Universal Robots URScript: test_first_drawing_6.script

def Machining1():
  # Default parameters:
  global speed_ms = 0.3
  global speed_rads = 0.75
  global accel_mss = 3
  global accel_radss = 1.2
  global blend_radius_m = 0.001

  # Add subprograms here
  # Start of main program
  # Program generated by RoboDK v5.6.5 for UR10e on 02/02/2024 17:00:01
  # Using nominal kinematics.
  blend_radius_m = 0.001
  speed_ms = 1.000
  # set_reference(p[0.133734, -0.230000, -0.011586, 0.000000, 0.000000, 0.000000])
  set_tcp(p[0.000000, 0.000000, 0.252000, 0.000000, 0.000000, 0.000000])
  # Show Tool
  movej([-0.330517, -0.652308, -2.595548, -1.464533, 1.570796, 1.240279],accel_radss,speed_rads,0,blend_radius_m)
  movel([-0.330517, -0.652308, -2.595548, -1.464533, 1.570796, 1.240279],accel_mss,speed_ms,0,blend_radius_m)
  # Splitting Linear movement in 6 (instruction 7: MoveL 3)
  movel([-0.330517, -0.658933, -2.623995, -1.429460, 1.570796, 1.240279],accel_mss,speed_ms,0,blend_radius_m)
  movel([-0.330517, -0.667915, -2.652250, -1.392224, 1.570796, 1.240279],accel_mss,speed_ms,0,blend_radius_m)
  movel([-0.330517, -0.679637, -2.680305, -1.352447, 1.570796, 1.240279],accel_mss,speed_ms,0,blend_radius_m)
  movel([-0.330517, -0.694570, -2.708148, -1.309671, 1.570796, 1.240279],accel_mss,speed_ms,0,blend_radius_m)
  movel([-0.330517, -0.713300, -2.735763, -1.263326, 1.570796, 1.240279],accel_mss,speed_ms,0,blend_radius_m)
  movel([-0.330517, -0.736556, -2.763126, -1.212708, 1.570796, 1.240279],accel_mss,speed_ms,0,blend_radius_m)
  movel([-0.330517, -0.736556, -2.763126, -1.212708, 1.570796, 1.240279],accel_mss,speed_ms,0,blend_radius_m)
  speed_ms = 1.000
  movel([-0.330517, -0.736556, -2.763126, -1.212708, 1.570796, 1.240279],accel_mss,speed_ms,0,blend_radius_m)
  movel([-0.330517, -0.736556, -2.763126, -1.212708, 1.570796, 1.240279],accel_mss,speed_ms,0,blend_radius_m)
  movel([-0.330517, -0.736556, -2.763126, -1.212708, 1.570796, 1.240279],accel_mss,speed_ms,0,blend_radius_m)
  speed_ms = 0.005
  movel([-0.330517, -0.709218, -2.730259, -1.272912, 1.570796, 1.240279],accel_mss,speed_ms,0,blend_radius_m)
  speed_ms = 1.000
  movel([-0.330517, -0.736556, -2.763126, -1.212708, 1.570796, 1.240279],accel_mss,speed_ms,0,blend_radius_m)
  speed_ms = 0.040
  movel([-0.330517, -0.736556, -2.763126, -1.212708, 1.570796, 1.240279],accel_mss,speed_ms,0,blend_radius_m)
  speed_ms = 1.000
  movel([-0.330517, -0.736556, -2.763126, -1.212708, 1.570796, 1.240279],accel_mss,speed_ms,0,blend_radius_m)
  # Splitting Linear movement in 8 (instruction 21: MoveL 12)
  movel([-0.265752, -0.726906, -2.764568, -1.220915, 1.570796, 1.305044],accel_mss,speed_ms,0,blend_radius_m)
  movel([-0.203429, -0.722340, -2.765235, -1.224814, 1.570796, 1.367367],accel_mss,speed_ms,0,blend_radius_m)
  movel([-0.144075, -0.722992, -2.765140, -1.224257, 1.570796, 1.426722],accel_mss,speed_ms,0,blend_radius_m)
  movel([-0.088098, -0.728842, -2.764283, -1.219264, 1.570796, 1.482698],accel_mss,speed_ms,0,blend_radius_m)
  movel([-0.035774, -0.739721, -2.762642, -1.210026, 1.570796, 1.535022],accel_mss,speed_ms,0,blend_radius_m)
  movel([0.012756, -0.755321, -2.760186, -1.196882, 1.570796, 1.583552],accel_mss,speed_ms,0,blend_radius_m)
  movel([0.057475, -0.775222, -2.756871, -1.180296, 1.570796, 1.628271],accel_mss,speed_ms,0,blend_radius_m)
  movel([0.098470, -0.798920, -2.752649, -1.160820, 1.570796, 1.669266],accel_mss,speed_ms,0,blend_radius_m)
  speed_ms = 0.005
  movel([0.098470, -0.837473, -2.784197, -1.090719, 1.570796, 1.669266],accel_mss,speed_ms,0,blend_radius_m)
  speed_ms = 0.025
  movel([0.094484, -0.848078, -2.782141, -1.082170, 1.570796, 1.665281],accel_mss,speed_ms,0,blend_radius_m)
  movel([0.092287, -0.853406, -2.781085, -1.077898, 1.570796, 1.663083],accel_mss,speed_ms,0,blend_radius_m)
  movel([0.089913, -0.858734, -2.780012, -1.073643, 1.570796, 1.660710],accel_mss,speed_ms,0,blend_radius_m)
  movel([0.087338, -0.864042, -2.778926, -1.069420, 1.570796, 1.658135],accel_mss,speed_ms,0,blend_radius_m)
  movel([0.084536, -0.869315, -2.777832, -1.065242, 1.570796, 1.655333],accel_mss,speed_ms,0,blend_radius_m)
  movel([0.081477, -0.874542, -2.776731, -1.061116, 1.570796, 1.652273],accel_mss,speed_ms,0,blend_radius_m)
  movel([0.078131, -0.879702, -2.775628, -1.057059, 1.570796, 1.648928],accel_mss,speed_ms,0,blend_radius_m)
  movel([0.079373, -0.877446, -2.776112, -1.058831, 1.570796, 1.650169],accel_mss,speed_ms,0,blend_radius_m)
  movel([0.080517, -0.874618, -2.776715, -1.061056, 1.570796, 1.651313],accel_mss,speed_ms,0,blend_radius_m)
  movel([0.081210, -0.871968, -2.777275, -1.063146, 1.570796, 1.652007],accel_mss,speed_ms,0,blend_radius_m)
  movel([0.081271, -0.870953, -2.777489, -1.063947, 1.570796, 1.652068],accel_mss,speed_ms,0,blend_radius_m)
  movel([0.081086, -0.870269, -2.777632, -1.064488, 1.570796, 1.651882],accel_mss,speed_ms,0,blend_radius_m)
  movel([0.080605, -0.869994, -2.777690, -1.064705, 1.570796, 1.651401],accel_mss,speed_ms,0,blend_radius_m)
  movel([0.079917, -0.870224, -2.777642, -1.064524, 1.570796, 1.650713],accel_mss,speed_ms,0,blend_radius_m)
  movel([0.079063, -0.870887, -2.777502, -1.063999, 1.570796, 1.649859],accel_mss,speed_ms,0,blend_radius_m)
  movel([0.078060, -0.871934, -2.777282, -1.063173, 1.570796, 1.648856],accel_mss,speed_ms,0,blend_radius_m)
  movel([0.075754, -0.874898, -2.776655, -1.060835, 1.570796, 1.646551],accel_mss,speed_ms,0,blend_radius_m)
  movel([0.073242, -0.878610, -2.775863, -1.057916, 1.570796, 1.644038],accel_mss,speed_ms,0,blend_radius_m)
  movel([0.068514, -0.886327, -2.774188, -1.051873, 1.570796, 1.639311],accel_mss,speed_ms,0,blend_radius_m)
  movel([0.065663, -0.891230, -2.773106, -1.048053, 1.570796, 1.636460],accel_mss,speed_ms,0,blend_radius_m)
  movel([0.061416, -0.898083, -2.771568, -1.042738, 1.570796, 1.632212],accel_mss,speed_ms,0,blend_radius_m)
  movel([0.059067, -0.901365, -2.770821, -1.040203, 1.570796, 1.629863],accel_mss,speed_ms,0,blend_radius_m)
  movel([0.056470, -0.904440, -2.770115, -1.037833, 1.570796, 1.627267],accel_mss,speed_ms,0,blend_radius_m)
  movel([0.057008, -0.903519, -2.770327, -1.038543, 1.570796, 1.627804],accel_mss,speed_ms,0,blend_radius_m)
  movel([0.057386, -0.902191, -2.770632, -1.039565, 1.570796, 1.628182],accel_mss,speed_ms,0,blend_radius_m)
  movel([0.057710, -0.898919, -2.771378, -1.042091, 1.570796, 1.628506],accel_mss,speed_ms,0,blend_radius_m)
  movel([0.057532, -0.895865, -2.772069, -1.044455, 1.570796, 1.628328],accel_mss,speed_ms,0,blend_radius_m)
  movel([0.057276, -0.894808, -2.772307, -1.045274, 1.570796, 1.628072],accel_mss,speed_ms,0,blend_radius_m)
  movel([0.056930, -0.894278, -2.772426, -1.045686, 1.570796, 1.627726],accel_mss,speed_ms,0,blend_radius_m)
  movel([0.055907, -0.894028, -2.772481, -1.045879, 1.570796, 1.626704],accel_mss,speed_ms,0,blend_radius_m)
  movel([0.054873, -0.894325, -2.772415, -1.045649, 1.570796, 1.625669],accel_mss,speed_ms,0,blend_radius_m)
  movel([0.053834, -0.895056, -2.772251, -1.045082, 1.570796, 1.624631],accel_mss,speed_ms,0,blend_radius_m)
  movel([0.052803, -0.896120, -2.772012, -1.044258, 1.570796, 1.623599],accel_mss,speed_ms,0,blend_radius_m)
  movel([0.050825, -0.898766, -2.771413, -1.042210, 1.570796, 1.621621],accel_mss,speed_ms,0,blend_radius_m)
  movel([0.049035, -0.901386, -2.770816, -1.040187, 1.570796, 1.619831],accel_mss,speed_ms,0,blend_radius_m)
  movel([0.046096, -0.905333, -2.769909, -1.037147, 1.570796, 1.616892],accel_mss,speed_ms,0,blend_radius_m)
  movel([0.043104, -0.908938, -2.769072, -1.034379, 1.570796, 1.613900],accel_mss,speed_ms,0,blend_radius_m)
  movel([0.039882, -0.912201, -2.768307, -1.031881, 1.570796, 1.610679],accel_mss,speed_ms,0,blend_radius_m)
  movel([0.036270, -0.915096, -2.767623, -1.029670, 1.570796, 1.607066],accel_mss,speed_ms,0,blend_radius_m)
  movel([0.038295, -0.912091, -2.768333, -1.031965, 1.570796, 1.609092],accel_mss,speed_ms,0,blend_radius_m)
  movel([0.039935, -0.909052, -2.769046, -1.034292, 1.570796, 1.610731],accel_mss,speed_ms,0,blend_radius_m)
  movel([0.040448, -0.907548, -2.769396, -1.035445, 1.570796, 1.611244],accel_mss,speed_ms,0,blend_radius_m)
  movel([0.040644, -0.906186, -2.769712, -1.036491, 1.570796, 1.611440],accel_mss,speed_ms,0,blend_radius_m)
  movel([0.040480, -0.905086, -2.769966, -1.037336, 1.570796, 1.611276],accel_mss,speed_ms,0,blend_radius_m)
  movel([0.039889, -0.904398, -2.770125, -1.037866, 1.570796, 1.610686],accel_mss,speed_ms,0,blend_radius_m)
  movel([0.038611, -0.904273, -2.770154, -1.037962, 1.570796, 1.609407],accel_mss,speed_ms,0,blend_radius_m)
  movel([0.036998, -0.904844, -2.770022, -1.037523, 1.570796, 1.607794],accel_mss,speed_ms,0,blend_radius_m)
  movel([0.035210, -0.905879, -2.769783, -1.036727, 1.570796, 1.606006],accel_mss,speed_ms,0,blend_radius_m)
  movel([0.033415, -0.907124, -2.769494, -1.035771, 1.570796, 1.604211],accel_mss,speed_ms,0,blend_radius_m)
  speed_ms = 0.005
  movel([0.033415, -0.898152, -2.763466, -1.050771, 1.570796, 1.604211],accel_mss,speed_ms,0,blend_radius_m)
  speed_ms = 0.040
  movel([0.037572, -0.930926, -2.755578, -1.025884, 1.570796, 1.608368],accel_mss,speed_ms,0,blend_radius_m)
  speed_ms = 0.005
  movel([0.037572, -0.940094, -2.761488, -1.010807, 1.570796, 1.608368],accel_mss,speed_ms,0,blend_radius_m)
  speed_ms = 0.025
  movel([0.038407, -0.937648, -2.762106, -1.012634, 1.570796, 1.609204],accel_mss,speed_ms,0,blend_radius_m)
  movel([0.039504, -0.935133, -2.762738, -1.014518, 1.570796, 1.610300],accel_mss,speed_ms,0,blend_radius_m)
  movel([0.040832, -0.932593, -2.763372, -1.016424, 1.570796, 1.611628],accel_mss,speed_ms,0,blend_radius_m)
  movel([0.042377, -0.930056, -2.764001, -1.018332, 1.570796, 1.613173],accel_mss,speed_ms,0,blend_radius_m)
  movel([0.044112, -0.927559, -2.764616, -1.020214, 1.570796, 1.614908],accel_mss,speed_ms,0,blend_radius_m)
  movel([0.046017, -0.925143, -2.765207, -1.022039, 1.570796, 1.616813],accel_mss,speed_ms,0,blend_radius_m)
  movel([0.048065, -0.922844, -2.765765, -1.023780, 1.570796, 1.618862],accel_mss,speed_ms,0,blend_radius_m)
  movel([0.050239, -0.920694, -2.766285, -1.025410, 1.570796, 1.621035],accel_mss,speed_ms,0,blend_radius_m)
  movel([0.053602, -0.917840, -2.766970, -1.027579, 1.570796, 1.624398],accel_mss,speed_ms,0,blend_radius_m)
  movel([0.056890, -0.915555, -2.767514, -1.029320, 1.570796, 1.627686],accel_mss,speed_ms,0,blend_radius_m)
  movel([0.060092, -0.913802, -2.767930, -1.030657, 1.570796, 1.630888],accel_mss,speed_ms,0,blend_radius_m)
  movel([0.063188, -0.912552, -2.768225, -1.031612, 1.570796, 1.633984],accel_mss,speed_ms,0,blend_radius_m)
  movel([0.066168, -0.911768, -2.768409, -1.032211, 1.570796, 1.636964],accel_mss,speed_ms,0,blend_radius_m)
  movel([0.069022, -0.911415, -2.768492, -1.032482, 1.570796, 1.639818],accel_mss,speed_ms,0,blend_radius_m)
  movel([0.071734, -0.911461, -2.768482, -1.032447, 1.570796, 1.642530],accel_mss,speed_ms,0,blend_radius_m)
  movel([0.074296, -0.911861, -2.768387, -1.032140, 1.570796, 1.645092],accel_mss,speed_ms,0,blend_radius_m)
  movel([0.076697, -0.912580, -2.768218, -1.031591, 1.570796, 1.647493],accel_mss,speed_ms,0,blend_radius_m)
  movel([0.078931, -0.913578, -2.767983, -1.030829, 1.570796, 1.649727],accel_mss,speed_ms,0,blend_radius_m)
  movel([0.082865, -0.916242, -2.767351, -1.028797, 1.570796, 1.653661],accel_mss,speed_ms,0,blend_radius_m)
  movel([0.086044, -0.919518, -2.766568, -1.026304, 1.570796, 1.656840],accel_mss,speed_ms,0,blend_radius_m)
  movel([0.088410, -0.923091, -2.765706, -1.023593, 1.570796, 1.659206],accel_mss,speed_ms,0,blend_radius_m)
  movel([0.090331, -0.927270, -2.764687, -1.020432, 1.570796, 1.661127],accel_mss,speed_ms,0,blend_radius_m)
  movel([0.091833, -0.931808, -2.763567, -1.017014, 1.570796, 1.662629],accel_mss,speed_ms,0,blend_radius_m)
  movel([0.092966, -0.936641, -2.762360, -1.013388, 1.570796, 1.663762],accel_mss,speed_ms,0,blend_radius_m)
  movel([0.093774, -0.941716, -2.761075, -1.009597, 1.570796, 1.664570],accel_mss,speed_ms,0,blend_radius_m)
  movel([0.094306, -0.946974, -2.759726, -1.005688, 1.570796, 1.665103],accel_mss,speed_ms,0,blend_radius_m)
  movel([0.094614, -0.952360, -2.758325, -1.001704, 1.570796, 1.665411],accel_mss,speed_ms,0,blend_radius_m)
  movel([0.094736, -0.963302, -2.755416, -0.993671, 1.570796, 1.665532],accel_mss,speed_ms,0,blend_radius_m)
  movel([0.094750, -0.970923, -2.753340, -0.988126, 1.570796, 1.665546],accel_mss,speed_ms,0,blend_radius_m)
  movel([0.095064, -0.974489, -2.752355, -0.985545, 1.570796, 1.665861],accel_mss,speed_ms,0,blend_radius_m)
  movel([0.095787, -0.977736, -2.751449, -0.983203, 1.570796, 1.666583],accel_mss,speed_ms,0,blend_radius_m)
  movel([0.097346, -0.981517, -2.750386, -0.980486, 1.570796, 1.668143],accel_mss,speed_ms,0,blend_radius_m)
  movel([0.098905, -0.985307, -2.749309, -0.977773, 1.570796, 1.669701],accel_mss,speed_ms,0,blend_radius_m)
  movel([0.099406, -0.987343, -2.748726, -0.976320, 1.570796, 1.670202],accel_mss,speed_ms,0,blend_radius_m)
  movel([0.099571, -0.989546, -2.748092, -0.974750, 1.570796, 1.670367],accel_mss,speed_ms,0,blend_radius_m)
  movel([0.099295, -0.991964, -2.747392, -0.973033, 1.570796, 1.670091],accel_mss,speed_ms,0,blend_radius_m)
  movel([0.098473, -0.994652, -2.746609, -0.971128, 1.570796, 1.669269],accel_mss,speed_ms,0,blend_radius_m)
  movel([0.101094, -0.987874, -2.748574, -0.975941, 1.570796, 1.671890],accel_mss,speed_ms,0,blend_radius_m)
  movel([0.103419, -0.981143, -2.750492, -0.980754, 1.570796, 1.674215],accel_mss,speed_ms,0,blend_radius_m)
  movel([0.107547, -0.967644, -2.754238, -0.990506, 1.570796, 1.678343],accel_mss,speed_ms,0,blend_radius_m)
  movel([0.109649, -0.960093, -2.756278, -0.996019, 1.570796, 1.680446],accel_mss,speed_ms,0,blend_radius_m)
  movel([0.111578, -0.952541, -2.758278, -1.001571, 1.570796, 1.682375],accel_mss,speed_ms,0,blend_radius_m)
  movel([0.115043, -0.937387, -2.762172, -1.012830, 1.570796, 1.685839],accel_mss,speed_ms,0,blend_radius_m)
  movel([0.118016, -0.922483, -2.765853, -1.024053, 1.570796, 1.688812],accel_mss,speed_ms,0,blend_radius_m)
  movel([0.119175, -0.915076, -2.767628, -1.029685, 1.570796, 1.689972],accel_mss,speed_ms,0,blend_radius_m)
  movel([0.119952, -0.907871, -2.769321, -1.035197, 1.570796, 1.690749],accel_mss,speed_ms,0,blend_radius_m)
  movel([0.120167, -0.902405, -2.770583, -1.039401, 1.570796, 1.690963],accel_mss,speed_ms,0,blend_radius_m)
  movel([0.120127, -0.897049, -2.771802, -1.043538, 1.570796, 1.690923],accel_mss,speed_ms,0,blend_radius_m)
  movel([0.120107, -0.891619, -2.773019, -1.047751, 1.570796, 1.690904],accel_mss,speed_ms,0,blend_radius_m)
  movel([0.120387, -0.885931, -2.774275, -1.052183, 1.570796, 1.691183],accel_mss,speed_ms,0,blend_radius_m)
  movel([0.120647, -0.884307, -2.774630, -1.053451, 1.570796, 1.691443],accel_mss,speed_ms,0,blend_radius_m)
  movel([0.121203, -0.882545, -2.775013, -1.054830, 1.570796, 1.692000],accel_mss,speed_ms,0,blend_radius_m)
  movel([0.122110, -0.880885, -2.775373, -1.056131, 1.570796, 1.692906],accel_mss,speed_ms,0,blend_radius_m)
  movel([0.122719, -0.880160, -2.775529, -1.056700, 1.570796, 1.693515],accel_mss,speed_ms,0,blend_radius_m)
  movel([0.123441, -0.879540, -2.775663, -1.057186, 1.570796, 1.694238],accel_mss,speed_ms,0,blend_radius_m)
  movel([0.124465, -0.879007, -2.775777, -1.057605, 1.570796, 1.695262],accel_mss,speed_ms,0,blend_radius_m)
  movel([0.125422, -0.878749, -2.775833, -1.057807, 1.570796, 1.696219],accel_mss,speed_ms,0,blend_radius_m)
  movel([0.130425, -0.878041, -2.775985, -1.058363, 1.570796, 1.701221],accel_mss,speed_ms,0,blend_radius_m)
  movel([0.134885, -0.878093, -2.775974, -1.058323, 1.570796, 1.705681],accel_mss,speed_ms,0,blend_radius_m)
  movel([0.138838, -0.878832, -2.775815, -1.057742, 1.570796, 1.709634],accel_mss,speed_ms,0,blend_radius_m)
  movel([0.142320, -0.880210, -2.775519, -1.056661, 1.570796, 1.713117],accel_mss,speed_ms,0,blend_radius_m)
  movel([0.145368, -0.882154, -2.775098, -1.055137, 1.570796, 1.716164],accel_mss,speed_ms,0,blend_radius_m)
  movel([0.148021, -0.884600, -2.774566, -1.053223, 1.570796, 1.718817],accel_mss,speed_ms,0,blend_radius_m)
  movel([0.150317, -0.887485, -2.773934, -1.050970, 1.570796, 1.721113],accel_mss,speed_ms,0,blend_radius_m)
  movel([0.152293, -0.890749, -2.773213, -1.048427, 1.570796, 1.723089],accel_mss,speed_ms,0,blend_radius_m)
  movel([0.153993, -0.894325, -2.772415, -1.045649, 1.570796, 1.724789],accel_mss,speed_ms,0,blend_radius_m)
  movel([0.155459, -0.898148, -2.771553, -1.042688, 1.570796, 1.726255],accel_mss,speed_ms,0,blend_radius_m)
  movel([0.157842, -0.906294, -2.769687, -1.036408, 1.570796, 1.728639],accel_mss,speed_ms,0,blend_radius_m)
  movel([0.161526, -0.922971, -2.765735, -1.023684, 1.570796, 1.732322],accel_mss,speed_ms,0,blend_radius_m)
  movel([0.162250, -0.925447, -2.765132, -1.021810, 1.570796, 1.733046],accel_mss,speed_ms,0,blend_radius_m)
  movel([0.162856, -0.926430, -2.764892, -1.021067, 1.570796, 1.733653],accel_mss,speed_ms,0,blend_radius_m)
  movel([0.163731, -0.927104, -2.764727, -1.020558, 1.570796, 1.734527],accel_mss,speed_ms,0,blend_radius_m)
  movel([0.165528, -0.927367, -2.764663, -1.020359, 1.570796, 1.736325],accel_mss,speed_ms,0,blend_radius_m)
  movel([0.166517, -0.927169, -2.764711, -1.020509, 1.570796, 1.737313],accel_mss,speed_ms,0,blend_radius_m)
  movel([0.167553, -0.926771, -2.764809, -1.020809, 1.570796, 1.738350],accel_mss,speed_ms,0,blend_radius_m)
  movel([0.169715, -0.925475, -2.765126, -1.021788, 1.570796, 1.740512],accel_mss,speed_ms,0,blend_radius_m)
  movel([0.171931, -0.923638, -2.765573, -1.023178, 1.570796, 1.742727],accel_mss,speed_ms,0,blend_radius_m)
  movel([0.174106, -0.921428, -2.766108, -1.024853, 1.570796, 1.744902],accel_mss,speed_ms,0,blend_radius_m)
  movel([0.176150, -0.919007, -2.766690, -1.026692, 1.570796, 1.746946],accel_mss,speed_ms,0,blend_radius_m)
  movel([0.177974, -0.916533, -2.767282, -1.028575, 1.570796, 1.748770],accel_mss,speed_ms,0,blend_radius_m)
  movel([0.179471, -0.914180, -2.767840, -1.030369, 1.570796, 1.750268],accel_mss,speed_ms,0,blend_radius_m)
  movel([0.181767, -0.910113, -2.768798, -1.033479, 1.570796, 1.752563],accel_mss,speed_ms,0,blend_radius_m)
  movel([0.183931, -0.905995, -2.769756, -1.036638, 1.570796, 1.754728],accel_mss,speed_ms,0,blend_radius_m)
  movel([0.187846, -0.897673, -2.771661, -1.043055, 1.570796, 1.758643],accel_mss,speed_ms,0,blend_radius_m)
  movel([0.191204, -0.889350, -2.773523, -1.049516, 1.570796, 1.762001],accel_mss,speed_ms,0,blend_radius_m)
  movel([0.193979, -0.881167, -2.775312, -1.055910, 1.570796, 1.764775],accel_mss,speed_ms,0,blend_radius_m)
  movel([0.194923, -0.878107, -2.775971, -1.058312, 1.570796, 1.765719],accel_mss,speed_ms,0,blend_radius_m)
  movel([0.196094, -0.874996, -2.776634, -1.060759, 1.570796, 1.766891],accel_mss,speed_ms,0,blend_radius_m)
  movel([0.196862, -0.873443, -2.776964, -1.061982, 1.570796, 1.767658],accel_mss,speed_ms,0,blend_radius_m)
  movel([0.197803, -0.871892, -2.777291, -1.063206, 1.570796, 1.768600],accel_mss,speed_ms,0,blend_radius_m)
  movel([0.198955, -0.870356, -2.777614, -1.064419, 1.570796, 1.769752],accel_mss,speed_ms,0,blend_radius_m)
  movel([0.200357, -0.868846, -2.777930, -1.065613, 1.570796, 1.771153],accel_mss,speed_ms,0,blend_radius_m)
  movel([0.202401, -0.867258, -2.778261, -1.066870, 1.570796, 1.773197],accel_mss,speed_ms,0,blend_radius_m)
  movel([0.204401, -0.866388, -2.778441, -1.067560, 1.570796, 1.775198],accel_mss,speed_ms,0,blend_radius_m)
  movel([0.206224, -0.866155, -2.778490, -1.067744, 1.570796, 1.777021],accel_mss,speed_ms,0,blend_radius_m)
  movel([0.207752, -0.866467, -2.778425, -1.067497, 1.570796, 1.778548],accel_mss,speed_ms,0,blend_radius_m)
  movel([0.209849, -0.867635, -2.778182, -1.066572, 1.570796, 1.780645],accel_mss,speed_ms,0,blend_radius_m)
  movel([0.211668, -0.869211, -2.777854, -1.065325, 1.570796, 1.782464],accel_mss,speed_ms,0,blend_radius_m)
  movel([0.214678, -0.873031, -2.777051, -1.062307, 1.570796, 1.785474],accel_mss,speed_ms,0,blend_radius_m)
  movel([0.215840, -0.875081, -2.776616, -1.060692, 1.570796, 1.786637],accel_mss,speed_ms,0,blend_radius_m)
  movel([0.216722, -0.877317, -2.776140, -1.058932, 1.570796, 1.787518],accel_mss,speed_ms,0,blend_radius_m)
  movel([0.217344, -0.879718, -2.775624, -1.057046, 1.570796, 1.788140],accel_mss,speed_ms,0,blend_radius_m)
  movel([0.217717, -0.882278, -2.775071, -1.055040, 1.570796, 1.788513],accel_mss,speed_ms,0,blend_radius_m)
  movel([0.217858, -0.884977, -2.774484, -1.052928, 1.570796, 1.788654],accel_mss,speed_ms,0,blend_radius_m)
  movel([0.217499, -0.890757, -2.773211, -1.048421, 1.570796, 1.788295],accel_mss,speed_ms,0,blend_radius_m)
  movel([0.217027, -0.893809, -2.772531, -1.046050, 1.570796, 1.787823],accel_mss,speed_ms,0,blend_radius_m)
  movel([0.215585, -0.900170, -2.771094, -1.041125, 1.570796, 1.786381],accel_mss,speed_ms,0,blend_radius_m)
  movel([0.213564, -0.906799, -2.769570, -1.036020, 1.570796, 1.784360],accel_mss,speed_ms,0,blend_radius_m)
  movel([0.211074, -0.913611, -2.767975, -1.030803, 1.570796, 1.781870],accel_mss,speed_ms,0,blend_radius_m)
  movel([0.208233, -0.920505, -2.766330, -1.025554, 1.570796, 1.779029],accel_mss,speed_ms,0,blend_radius_m)
  movel([0.203631, -0.930571, -2.763874, -1.017944, 1.570796, 1.774427],accel_mss,speed_ms,0,blend_radius_m)
  movel([0.201108, -0.935588, -2.762624, -1.014176, 1.570796, 1.771904],accel_mss,speed_ms,0,blend_radius_m)
  movel([0.198410, -0.940566, -2.761368, -1.010455, 1.570796, 1.769207],accel_mss,speed_ms,0,blend_radius_m)
  movel([0.195524, -0.945474, -2.760113, -1.006802, 1.570796, 1.766320],accel_mss,speed_ms,0,blend_radius_m)
  movel([0.192436, -0.950291, -2.758866, -1.003232, 1.570796, 1.763232],accel_mss,speed_ms,0,blend_radius_m)
  movel([0.189119, -0.955003, -2.757630, -0.999756, 1.570796, 1.759915],accel_mss,speed_ms,0,blend_radius_m)
  movel([0.185564, -0.959579, -2.756415, -0.996395, 1.570796, 1.756360],accel_mss,speed_ms,0,blend_radius_m)
  movel([0.180277, -0.965730, -2.754759, -0.991900, 1.570796, 1.751073],accel_mss,speed_ms,0,blend_radius_m)
  movel([0.177371, -0.968805, -2.753921, -0.989663, 1.570796, 1.748167],accel_mss,speed_ms,0,blend_radius_m)
  movel([0.174357, -0.971712, -2.753123, -0.987554, 1.570796, 1.745154],accel_mss,speed_ms,0,blend_radius_m)
  movel([0.171294, -0.974326, -2.752400, -0.985663, 1.570796, 1.742090],accel_mss,speed_ms,0,blend_radius_m)
  movel([0.168232, -0.976525, -2.751788, -0.984076, 1.570796, 1.739028],accel_mss,speed_ms,0,blend_radius_m)
  movel([0.165220, -0.978184, -2.751324, -0.982881, 1.570796, 1.736016],accel_mss,speed_ms,0,blend_radius_m)
  movel([0.163750, -0.978776, -2.751158, -0.982455, 1.570796, 1.734546],accel_mss,speed_ms,0,blend_radius_m)
  movel([0.162314, -0.979184, -2.751043, -0.982162, 1.570796, 1.733110],accel_mss,speed_ms,0,blend_radius_m)
  movel([0.160767, -0.979407, -2.750981, -0.982001, 1.570796, 1.731564],accel_mss,speed_ms,0,blend_radius_m)
  movel([0.159366, -0.979372, -2.750991, -0.982027, 1.570796, 1.730163],accel_mss,speed_ms,0,blend_radius_m)
  movel([0.158098, -0.979106, -2.751065, -0.982218, 1.570796, 1.728894],accel_mss,speed_ms,0,blend_radius_m)
  movel([0.156956, -0.978625, -2.751200, -0.982563, 1.570796, 1.727752],accel_mss,speed_ms,0,blend_radius_m)
  movel([0.155007, -0.977127, -2.751620, -0.983642, 1.570796, 1.725804],accel_mss,speed_ms,0,blend_radius_m)
  movel([0.153455, -0.975052, -2.752199, -0.985139, 1.570796, 1.724251],accel_mss,speed_ms,0,blend_radius_m)
  movel([0.152226, -0.972588, -2.752881, -0.986920, 1.570796, 1.723022],accel_mss,speed_ms,0,blend_radius_m)
  movel([0.151254, -0.969917, -2.753617, -0.988856, 1.570796, 1.722051],accel_mss,speed_ms,0,blend_radius_m)
  movel([0.149812, -0.964692, -2.755040, -0.992657, 1.570796, 1.720608],accel_mss,speed_ms,0,blend_radius_m)
  movel([0.149169, -0.962231, -2.755704, -0.994453, 1.570796, 1.719965],accel_mss,speed_ms,0,blend_radius_m)
  movel([0.148254, -0.960029, -2.756295, -0.996065, 1.570796, 1.719050],accel_mss,speed_ms,0,blend_radius_m)
  movel([0.147575, -0.959185, -2.756520, -0.996684, 1.570796, 1.718371],accel_mss,speed_ms,0,blend_radius_m)
  movel([0.146683, -0.958596, -2.756677, -0.997116, 1.570796, 1.717479],accel_mss,speed_ms,0,blend_radius_m)
  movel([0.145535, -0.958328, -2.756749, -0.997313, 1.570796, 1.716332],accel_mss,speed_ms,0,blend_radius_m)
  movel([0.144083, -0.958440, -2.756719, -0.997230, 1.570796, 1.714879],accel_mss,speed_ms,0,blend_radius_m)
  movel([0.144394, -0.958486, -2.756707, -0.997197, 1.570796, 1.715191],accel_mss,speed_ms,0,blend_radius_m)
  movel([0.144561, -0.958767, -2.756632, -0.996990, 1.570796, 1.715357],accel_mss,speed_ms,0,blend_radius_m)
  movel([0.144480, -0.959980, -2.756308, -0.996101, 1.570796, 1.715276],accel_mss,speed_ms,0,blend_radius_m)
  movel([0.143903, -0.961959, -2.755777, -0.994652, 1.570796, 1.714700],accel_mss,speed_ms,0,blend_radius_m)
  movel([0.142911, -0.964578, -2.755071, -0.992740, 1.570796, 1.713708],accel_mss,speed_ms,0,blend_radius_m)
  movel([0.139967, -0.971238, -2.753254, -0.987898, 1.570796, 1.710763],accel_mss,speed_ms,0,blend_radius_m)
  movel([0.136215, -0.978975, -2.751102, -0.982312, 1.570796, 1.707011],accel_mss,speed_ms,0,blend_radius_m)
  movel([0.128486, -0.993946, -2.746815, -0.971628, 1.570796, 1.699282],accel_mss,speed_ms,0,blend_radius_m)
  movel([0.123866, -1.002374, -2.744329, -0.965686, 1.570796, 1.694663],accel_mss,speed_ms,0,blend_radius_m)
  movel([0.118500, -1.011014, -2.741724, -0.959651, 1.570796, 1.689296],accel_mss,speed_ms,0,blend_radius_m)
  movel([0.113088, -1.019425, -2.739133, -0.953832, 1.570796, 1.683885],accel_mss,speed_ms,0,blend_radius_m)
  movel([0.107607, -1.027694, -2.736531, -0.948164, 1.570796, 1.678403],accel_mss,speed_ms,0,blend_radius_m)
  movel([0.096784, -1.043415, -2.731434, -0.937539, 1.570796, 1.667580],accel_mss,speed_ms,0,blend_radius_m)
  movel([0.091340, -1.050721, -2.728997, -0.932671, 1.570796, 1.662136],accel_mss,speed_ms,0,blend_radius_m)
  movel([0.088492, -1.054219, -2.727815, -0.930356, 1.570796, 1.659288],accel_mss,speed_ms,0,blend_radius_m)
  movel([0.085541, -1.057575, -2.726671, -0.928144, 1.570796, 1.656337],accel_mss,speed_ms,0,blend_radius_m)
  movel([0.082458, -1.060760, -2.725576, -0.926053, 1.570796, 1.653255],accel_mss,speed_ms,0,blend_radius_m)
  movel([0.079236, -1.063748, -2.724541, -0.924100, 1.570796, 1.650032],accel_mss,speed_ms,0,blend_radius_m)
  movel([0.080076, -1.057742, -2.726613, -0.928034, 1.570796, 1.650872],accel_mss,speed_ms,0,blend_radius_m)
  movel([0.080087, -1.056070, -2.727185, -0.929134, 1.570796, 1.650884],accel_mss,speed_ms,0,blend_radius_m)
  movel([0.079804, -1.055496, -2.727380, -0.929512, 1.570796, 1.650600],accel_mss,speed_ms,0,blend_radius_m)
  movel([0.079211, -1.055294, -2.727449, -0.929646, 1.570796, 1.650008],accel_mss,speed_ms,0,blend_radius_m)
  movel([0.078545, -1.055474, -2.727388, -0.929527, 1.570796, 1.649341],accel_mss,speed_ms,0,blend_radius_m)
  movel([0.077831, -1.055896, -2.727244, -0.929249, 1.570796, 1.648627],accel_mss,speed_ms,0,blend_radius_m)
  movel([0.074420, -1.058581, -2.726326, -0.927482, 1.570796, 1.645216],accel_mss,speed_ms,0,blend_radius_m)
  movel([0.072411, -1.059837, -2.725894, -0.926658, 1.570796, 1.643207],accel_mss,speed_ms,0,blend_radius_m)
  movel([0.070406, -1.060807, -2.725560, -0.926022, 1.570796, 1.641202],accel_mss,speed_ms,0,blend_radius_m)
  movel([0.068457, -1.061467, -2.725331, -0.925590, 1.570796, 1.639253],accel_mss,speed_ms,0,blend_radius_m)
  movel([0.067876, -1.061499, -2.725320, -0.925569, 1.570796, 1.638673],accel_mss,speed_ms,0,blend_radius_m)
  movel([0.067717, -1.061162, -2.725437, -0.925790, 1.570796, 1.638514],accel_mss,speed_ms,0,blend_radius_m)
  movel([0.068293, -1.059355, -2.726060, -0.926974, 1.570796, 1.639089],accel_mss,speed_ms,0,blend_radius_m)
  movel([0.068248, -1.058832, -2.726239, -0.927317, 1.570796, 1.639044],accel_mss,speed_ms,0,blend_radius_m)
  movel([0.067937, -1.058525, -2.726345, -0.927519, 1.570796, 1.638733],accel_mss,speed_ms,0,blend_radius_m)
  movel([0.067444, -1.058429, -2.726378, -0.927582, 1.570796, 1.638240],accel_mss,speed_ms,0,blend_radius_m)
  movel([0.066848, -1.058544, -2.726338, -0.927507, 1.570796, 1.637644],accel_mss,speed_ms,0,blend_radius_m)
  movel([0.065582, -1.059240, -2.726099, -0.927049, 1.570796, 1.636378],accel_mss,speed_ms,0,blend_radius_m)
  movel([0.056656, -1.066547, -2.723565, -0.922277, 1.570796, 1.627452],accel_mss,speed_ms,0,blend_radius_m)
  movel([0.059293, -1.063911, -2.724484, -0.923994, 1.570796, 1.630089],accel_mss,speed_ms,0,blend_radius_m)
  movel([0.061894, -1.061075, -2.725467, -0.925847, 1.570796, 1.632691],accel_mss,speed_ms,0,blend_radius_m)
  movel([0.064438, -1.058090, -2.726494, -0.927805, 1.570796, 1.635234],accel_mss,speed_ms,0,blend_radius_m)
  movel([0.066915, -1.054985, -2.727555, -0.929850, 1.570796, 1.637712],accel_mss,speed_ms,0,blend_radius_m)
  movel([0.071603, -1.048575, -2.729718, -0.934097, 1.570796, 1.642399],accel_mss,speed_ms,0,blend_radius_m)
  movel([0.075821, -1.042175, -2.731844, -0.938370, 1.570796, 1.646617],accel_mss,speed_ms,0,blend_radius_m)
  movel([0.080132, -1.035147, -2.734140, -0.943102, 1.570796, 1.650928],accel_mss,speed_ms,0,blend_radius_m)
  movel([0.084250, -1.027966, -2.736445, -0.947978, 1.570796, 1.655047],accel_mss,speed_ms,0,blend_radius_m)
  movel([0.086168, -1.024338, -2.737594, -0.950458, 1.570796, 1.656965],accel_mss,speed_ms,0,blend_radius_m)
  movel([0.087963, -1.020694, -2.738737, -0.952958, 1.570796, 1.658760],accel_mss,speed_ms,0,blend_radius_m)
  movel([0.089601, -1.017048, -2.739870, -0.955470, 1.570796, 1.660397],accel_mss,speed_ms,0,blend_radius_m)
  movel([0.091057, -1.013402, -2.740994, -0.957993, 1.570796, 1.661853],accel_mss,speed_ms,0,blend_radius_m)
  movel([0.091816, -1.011152, -2.741682, -0.959555, 1.570796, 1.662613],accel_mss,speed_ms,0,blend_radius_m)
  movel([0.092410, -1.008926, -2.742359, -0.961105, 1.570796, 1.663206],accel_mss,speed_ms,0,blend_radius_m)
  movel([0.093141, -1.004571, -2.743672, -0.964146, 1.570796, 1.663937],accel_mss,speed_ms,0,blend_radius_m)
  movel([0.093305, -1.000395, -2.744917, -0.967076, 1.570796, 1.664101],accel_mss,speed_ms,0,blend_radius_m)
  movel([0.092955, -0.996450, -2.746082, -0.969857, 1.570796, 1.663751],accel_mss,speed_ms,0,blend_radius_m)
  movel([0.092159, -0.992782, -2.747155, -0.972453, 1.570796, 1.662955],accel_mss,speed_ms,0,blend_radius_m)
  movel([0.090980, -0.989443, -2.748122, -0.974824, 1.570796, 1.661776],accel_mss,speed_ms,0,blend_radius_m)
  movel([0.089473, -0.986490, -2.748971, -0.976928, 1.570796, 1.660269],accel_mss,speed_ms,0,blend_radius_m)
  movel([0.087711, -0.983965, -2.749691, -0.978732, 1.570796, 1.658507],accel_mss,speed_ms,0,blend_radius_m)
  movel([0.086357, -0.982932, -2.749985, -0.979472, 1.570796, 1.657154],accel_mss,speed_ms,0,blend_radius_m)
  movel([0.084665, -0.982603, -2.750078, -0.979707, 1.570796, 1.655461],accel_mss,speed_ms,0,blend_radius_m)
  movel([0.082738, -0.982926, -2.749987, -0.979476, 1.570796, 1.653534],accel_mss,speed_ms,0,blend_radius_m)
  movel([0.080685, -0.983843, -2.749726, -0.978819, 1.570796, 1.651481],accel_mss,speed_ms,0,blend_radius_m)
  movel([0.078604, -0.985294, -2.749313, -0.977782, 1.570796, 1.649400],accel_mss,speed_ms,0,blend_radius_m)
  movel([0.076600, -0.987221, -2.748761, -0.976406, 1.570796, 1.647396],accel_mss,speed_ms,0,blend_radius_m)
  movel([0.074785, -0.989556, -2.748089, -0.974743, 1.570796, 1.645582],accel_mss,speed_ms,0,blend_radius_m)
  movel([0.073255, -0.992240, -2.747312, -0.972837, 1.570796, 1.644052],accel_mss,speed_ms,0,blend_radius_m)
  movel([0.071220, -0.996348, -2.746112, -0.969929, 1.570796, 1.642016],accel_mss,speed_ms,0,blend_radius_m)
  movel([0.069032, -1.000411, -2.744913, -0.967065, 1.570796, 1.639828],accel_mss,speed_ms,0,blend_radius_m)
  movel([0.066672, -1.004395, -2.743725, -0.964270, 1.570796, 1.637469],accel_mss,speed_ms,0,blend_radius_m)
  movel([0.064115, -1.008273, -2.742556, -0.961559, 1.570796, 1.634912],accel_mss,speed_ms,0,blend_radius_m)
  movel([0.061349, -1.012012, -2.741419, -0.958958, 1.570796, 1.632145],accel_mss,speed_ms,0,blend_radius_m)
  movel([0.058346, -1.015587, -2.740322, -0.956480, 1.570796, 1.629142],accel_mss,speed_ms,0,blend_radius_m)
  movel([0.055086, -1.018973, -2.739273, -0.954143, 1.570796, 1.625883],accel_mss,speed_ms,0,blend_radius_m)
  movel([0.051553, -1.022140, -2.738285, -0.951965, 1.570796, 1.622350],accel_mss,speed_ms,0,blend_radius_m)
  movel([0.049638, -1.023581, -2.737832, -0.950976, 1.570796, 1.620435],accel_mss,speed_ms,0,blend_radius_m)
  movel([0.047695, -1.024799, -2.737448, -0.950142, 1.570796, 1.618491],accel_mss,speed_ms,0,blend_radius_m)
  movel([0.043791, -1.026823, -2.736808, -0.948758, 1.570796, 1.614588],accel_mss,speed_ms,0,blend_radius_m)
  movel([0.040756, -1.028106, -2.736400, -0.947883, 1.570796, 1.611552],accel_mss,speed_ms,0,blend_radius_m)
  movel([0.037886, -1.028957, -2.736129, -0.947303, 1.570796, 1.608683],accel_mss,speed_ms,0,blend_radius_m)
  movel([0.035183, -1.029408, -2.735985, -0.946996, 1.570796, 1.605979],accel_mss,speed_ms,0,blend_radius_m)
  movel([0.032632, -1.029495, -2.735958, -0.946937, 1.570796, 1.603429],accel_mss,speed_ms,0,blend_radius_m)
  movel([0.030229, -1.029253, -2.736035, -0.947101, 1.570796, 1.601025],accel_mss,speed_ms,0,blend_radius_m)
  movel([0.027965, -1.028713, -2.736207, -0.947469, 1.570796, 1.598761],accel_mss,speed_ms,0,blend_radius_m)
  movel([0.025843, -1.027903, -2.736465, -0.948021, 1.570796, 1.596639],accel_mss,speed_ms,0,blend_radius_m)
  movel([0.023853, -1.026860, -2.736796, -0.948733, 1.570796, 1.594650],accel_mss,speed_ms,0,blend_radius_m)
  movel([0.021991, -1.025616, -2.737190, -0.949583, 1.570796, 1.592787],accel_mss,speed_ms,0,blend_radius_m)
  movel([0.020254, -1.024192, -2.737640, -0.950557, 1.570796, 1.591051],accel_mss,speed_ms,0,blend_radius_m)
  movel([0.017143, -1.020959, -2.738654, -0.952776, 1.570796, 1.587940],accel_mss,speed_ms,0,blend_radius_m)
  movel([0.014492, -1.017403, -2.739761, -0.955225, 1.570796, 1.585288],accel_mss,speed_ms,0,blend_radius_m)
  movel([0.012279, -1.013785, -2.740876, -0.957728, 1.570796, 1.583076],accel_mss,speed_ms,0,blend_radius_m)
  movel([0.010780, -1.010844, -2.741776, -0.959769, 1.570796, 1.581576],accel_mss,speed_ms,0,blend_radius_m)
  movel([0.009435, -1.007642, -2.742747, -0.961999, 1.570796, 1.580232],accel_mss,speed_ms,0,blend_radius_m)
  movel([0.008265, -1.004187, -2.743787, -0.964415, 1.570796, 1.579062],accel_mss,speed_ms,0,blend_radius_m)
  movel([0.007306, -1.000492, -2.744889, -0.967009, 1.570796, 1.578102],accel_mss,speed_ms,0,blend_radius_m)
  movel([0.006575, -0.996570, -2.746047, -0.969772, 1.570796, 1.577371],accel_mss,speed_ms,0,blend_radius_m)
  movel([0.006105, -0.992433, -2.747256, -0.972700, 1.570796, 1.576901],accel_mss,speed_ms,0,blend_radius_m)
  movel([0.005928, -0.988091, -2.748512, -0.975787, 1.570796, 1.576724],accel_mss,speed_ms,0,blend_radius_m)
  movel([0.006071, -0.983555, -2.749808, -0.979026, 1.570796, 1.576868],accel_mss,speed_ms,0,blend_radius_m)
  movel([0.006563, -0.978834, -2.751142, -0.982413, 1.570796, 1.577359],accel_mss,speed_ms,0,blend_radius_m)
  movel([0.007436, -0.973949, -2.752505, -0.985935, 1.570796, 1.578232],accel_mss,speed_ms,0,blend_radius_m)
  movel([0.008720, -0.968900, -2.753895, -0.989593, 1.570796, 1.579516],accel_mss,speed_ms,0,blend_radius_m)
  movel([0.010453, -0.963704, -2.755308, -0.993378, 1.570796, 1.581249],accel_mss,speed_ms,0,blend_radius_m)
  movel([0.012661, -0.958375, -2.756736, -0.997278, 1.570796, 1.583458],accel_mss,speed_ms,0,blend_radius_m)
  movel([0.015384, -0.952920, -2.758178, -1.001291, 1.570796, 1.586181],accel_mss,speed_ms,0,blend_radius_m)
  movel([0.018649, -0.947365, -2.759625, -1.005399, 1.570796, 1.589446],accel_mss,speed_ms,0,blend_radius_m)
  movel([0.022491, -0.941719, -2.761075, -1.009595, 1.570796, 1.593287],accel_mss,speed_ms,0,blend_radius_m)
  movel([0.024161, -0.939594, -2.761615, -1.011180, 1.570796, 1.594957],accel_mss,speed_ms,0,blend_radius_m)
  movel([0.025079, -0.938637, -2.761857, -1.011895, 1.570796, 1.595875],accel_mss,speed_ms,0,blend_radius_m)
  movel([0.026054, -0.937835, -2.762059, -1.012495, 1.570796, 1.596851],accel_mss,speed_ms,0,blend_radius_m)
  movel([0.027520, -0.937088, -2.762248, -1.013054, 1.570796, 1.598316],accel_mss,speed_ms,0,blend_radius_m)
  movel([0.028823, -0.936912, -2.762292, -1.013185, 1.570796, 1.599619],accel_mss,speed_ms,0,blend_radius_m)
  movel([0.029911, -0.937209, -2.762217, -1.012963, 1.570796, 1.600707],accel_mss,speed_ms,0,blend_radius_m)
  movel([0.030731, -0.937876, -2.762049, -1.012464, 1.570796, 1.601527],accel_mss,speed_ms,0,blend_radius_m)
  movel([0.031881, -0.940032, -2.761504, -1.010853, 1.570796, 1.602677],accel_mss,speed_ms,0,blend_radius_m)
  movel([0.032501, -0.942703, -2.760824, -1.008862, 1.570796, 1.603297],accel_mss,speed_ms,0,blend_radius_m)
  movel([0.033157, -0.948460, -2.759342, -1.004587, 1.570796, 1.603954],accel_mss,speed_ms,0,blend_radius_m)
  movel([0.033560, -0.949351, -2.759110, -1.003928, 1.570796, 1.604356],accel_mss,speed_ms,0,blend_radius_m)
  movel([0.034009, -0.949386, -2.759101, -1.003902, 1.570796, 1.604805],accel_mss,speed_ms,0,blend_radius_m)
  movel([0.034702, -0.949062, -2.759186, -1.004142, 1.570796, 1.605499],accel_mss,speed_ms,0,blend_radius_m)
  movel([0.035843, -0.946344, -2.759889, -1.006156, 1.570796, 1.606639],accel_mss,speed_ms,0,blend_radius_m)
  movel([0.036834, -0.943600, -2.760594, -1.008195, 1.570796, 1.607630],accel_mss,speed_ms,0,blend_radius_m)
  movel([0.037444, -0.952233, -2.758358, -1.001798, 1.570796, 1.608241],accel_mss,speed_ms,0,blend_radius_m)
  movel([0.038358, -0.960568, -2.756151, -0.995670, 1.570796, 1.609155],accel_mss,speed_ms,0,blend_radius_m)
  movel([0.039568, -0.968608, -2.753975, -0.989806, 1.570796, 1.610365],accel_mss,speed_ms,0,blend_radius_m)
  movel([0.041067, -0.976361, -2.751834, -0.984194, 1.570796, 1.611863],accel_mss,speed_ms,0,blend_radius_m)
  movel([0.041844, -0.979624, -2.750920, -0.981845, 1.570796, 1.612640],accel_mss,speed_ms,0,blend_radius_m)
  movel([0.042968, -0.982777, -2.750029, -0.979583, 1.570796, 1.613764],accel_mss,speed_ms,0,blend_radius_m)
  movel([0.043724, -0.984173, -2.749632, -0.978584, 1.570796, 1.614520],accel_mss,speed_ms,0,blend_radius_m)
  movel([0.044642, -0.985370, -2.749291, -0.977728, 1.570796, 1.615439],accel_mss,speed_ms,0,blend_radius_m)
  movel([0.045753, -0.986310, -2.749022, -0.977056, 1.570796, 1.616549],accel_mss,speed_ms,0,blend_radius_m)
  movel([0.047082, -0.986935, -2.748843, -0.976610, 1.570796, 1.617878],accel_mss,speed_ms,0,blend_radius_m)
  movel([0.048145, -0.987141, -2.748784, -0.976464, 1.570796, 1.618941],accel_mss,speed_ms,0,blend_radius_m)
  movel([0.050510, -0.986919, -2.748848, -0.976622, 1.570796, 1.621306],accel_mss,speed_ms,0,blend_radius_m)
  movel([0.051789, -0.986524, -2.748961, -0.976904, 1.570796, 1.622585],accel_mss,speed_ms,0,blend_radius_m)
  movel([0.054481, -0.985253, -2.749325, -0.977811, 1.570796, 1.625277],accel_mss,speed_ms,0,blend_radius_m)
  movel([0.057280, -0.983439, -2.749841, -0.979109, 1.570796, 1.628077],accel_mss,speed_ms,0,blend_radius_m)
  movel([0.060093, -0.981218, -2.750470, -0.980701, 1.570796, 1.630889],accel_mss,speed_ms,0,blend_radius_m)
  movel([0.062827, -0.978710, -2.751177, -0.982503, 1.570796, 1.633623],accel_mss,speed_ms,0,blend_radius_m)
  movel([0.065387, -0.976051, -2.751920, -0.984418, 1.570796, 1.636184],accel_mss,speed_ms,0,blend_radius_m)
  movel([0.067670, -0.973373, -2.752664, -0.986352, 1.570796, 1.638466],accel_mss,speed_ms,0,blend_radius_m)
  speed_ms = 0.005
  movel([0.067670, -0.964047, -2.746880, -1.001462, 1.570796, 1.638466],accel_mss,speed_ms,0,blend_radius_m)
  speed_ms = 0.040
  movel([0.054777, -0.972239, -2.744611, -0.995539, 1.570796, 1.625574],accel_mss,speed_ms,0,blend_radius_m)
  speed_ms = 0.005
  movel([0.054777, -0.981598, -2.750363, -0.980428, 1.570796, 1.625574],accel_mss,speed_ms,0,blend_radius_m)
  speed_ms = 0.025
  movel([0.056594, -0.979364, -2.750993, -0.982032, 1.570796, 1.627391],accel_mss,speed_ms,0,blend_radius_m)
  movel([0.060089, -0.974446, -2.752367, -0.985576, 1.570796, 1.630885],accel_mss,speed_ms,0,blend_radius_m)
  movel([0.061733, -0.971814, -2.753095, -0.987480, 1.570796, 1.632530],accel_mss,speed_ms,0,blend_radius_m)
  movel([0.064740, -0.966337, -2.754594, -0.991458, 1.570796, 1.635536],accel_mss,speed_ms,0,blend_radius_m)
  movel([0.067277, -0.960747, -2.756103, -0.995539, 1.570796, 1.638073],accel_mss,speed_ms,0,blend_radius_m)
  movel([0.068328, -0.957982, -2.756841, -0.997566, 1.570796, 1.639124],accel_mss,speed_ms,0,blend_radius_m)
  movel([0.069210, -0.955271, -2.757559, -0.999559, 1.570796, 1.640006],accel_mss,speed_ms,0,blend_radius_m)
  movel([0.070403, -0.950139, -2.758905, -1.003345, 1.570796, 1.641199],accel_mss,speed_ms,0,blend_radius_m)
  movel([0.070684, -0.947770, -2.759520, -1.005098, 1.570796, 1.641480],accel_mss,speed_ms,0,blend_radius_m)
  movel([0.070726, -0.945583, -2.760085, -1.006721, 1.570796, 1.641522],accel_mss,speed_ms,0,blend_radius_m)
  movel([0.070518, -0.943600, -2.760594, -1.008195, 1.570796, 1.641314],accel_mss,speed_ms,0,blend_radius_m)
  movel([0.070039, -0.941852, -2.761041, -1.009496, 1.570796, 1.640836],accel_mss,speed_ms,0,blend_radius_m)
  movel([0.069145, -0.939957, -2.761523, -1.010910, 1.570796, 1.639941],accel_mss,speed_ms,0,blend_radius_m)
  movel([0.067993, -0.938333, -2.761934, -1.012122, 1.570796, 1.638790],accel_mss,speed_ms,0,blend_radius_m)
  movel([0.066567, -0.937058, -2.762255, -1.013076, 1.570796, 1.637363],accel_mss,speed_ms,0,blend_radius_m)
  movel([0.064853, -0.936213, -2.762468, -1.013709, 1.570796, 1.635649],accel_mss,speed_ms,0,blend_radius_m)
  movel([0.062833, -0.935875, -2.762552, -1.013962, 1.570796, 1.633630],accel_mss,speed_ms,0,blend_radius_m)
  movel([0.060502, -0.936120, -2.762491, -1.013778, 1.570796, 1.631299],accel_mss,speed_ms,0,blend_radius_m)
  movel([0.057846, -0.937027, -2.762263, -1.013099, 1.570796, 1.628642],accel_mss,speed_ms,0,blend_radius_m)
  movel([0.054857, -0.938658, -2.761851, -1.011879, 1.570796, 1.625654],accel_mss,speed_ms,0,blend_radius_m)
  movel([0.052795, -0.940155, -2.761472, -1.010761, 1.570796, 1.623592],accel_mss,speed_ms,0,blend_radius_m)
  movel([0.050789, -0.941944, -2.761017, -1.009428, 1.570796, 1.621585],accel_mss,speed_ms,0,blend_radius_m)
  movel([0.048907, -0.943948, -2.760505, -1.007936, 1.570796, 1.619703],accel_mss,speed_ms,0,blend_radius_m)
  movel([0.047206, -0.946097, -2.759953, -1.006339, 1.570796, 1.618002],accel_mss,speed_ms,0,blend_radius_m)
  movel([0.045744, -0.948321, -2.759378, -1.004690, 1.570796, 1.616540],accel_mss,speed_ms,0,blend_radius_m)
  movel([0.044580, -0.950550, -2.758798, -1.003041, 1.570796, 1.615376],accel_mss,speed_ms,0,blend_radius_m)
  movel([0.043774, -0.952714, -2.758232, -1.001443, 1.570796, 1.614571],accel_mss,speed_ms,0,blend_radius_m)
  movel([0.043376, -0.954750, -2.757697, -0.999942, 1.570796, 1.614172],accel_mss,speed_ms,0,blend_radius_m)
  speed_ms = 0.005
  movel([0.043376, -0.945508, -2.751842, -1.015040, 1.570796, 1.614172],accel_mss,speed_ms,0,blend_radius_m)
  speed_ms = 0.040
  # Splitting Linear movement in 2 (instruction 399: MoveL 378)
  movel([0.095251, -0.952183, -2.750083, -1.010123, 1.570796, 1.666048],accel_mss,speed_ms,0,blend_radius_m)
  movel([0.144369, -0.962810, -2.747219, -1.002360, 1.570796, 1.715166],accel_mss,speed_ms,0,blend_radius_m)
  speed_ms = 0.005
  movel([0.144369, -0.972131, -2.753008, -0.987251, 1.570796, 1.715166],accel_mss,speed_ms,0,blend_radius_m)
  speed_ms = 0.025
  movel([0.142576, -0.982664, -2.750061, -0.979664, 1.570796, 1.713373],accel_mss,speed_ms,0,blend_radius_m)
  movel([0.141323, -0.988007, -2.748536, -0.975846, 1.570796, 1.712119],accel_mss,speed_ms,0,blend_radius_m)
  movel([0.140478, -0.990766, -2.747740, -0.973883, 1.570796, 1.711274],accel_mss,speed_ms,0,blend_radius_m)
  movel([0.139439, -0.993604, -2.746915, -0.971870, 1.570796, 1.710235],accel_mss,speed_ms,0,blend_radius_m)
  movel([0.138085, -0.996654, -2.746022, -0.969712, 1.570796, 1.708881],accel_mss,speed_ms,0,blend_radius_m)
  movel([0.137248, -0.998165, -2.745577, -0.968647, 1.570796, 1.708044],accel_mss,speed_ms,0,blend_radius_m)
  movel([0.136253, -0.999641, -2.745141, -0.967607, 1.570796, 1.707050],accel_mss,speed_ms,0,blend_radius_m)
  movel([0.136298, -0.997342, -2.745820, -0.969227, 1.570796, 1.707094],accel_mss,speed_ms,0,blend_radius_m)
  movel([0.135952, -0.995298, -2.746420, -0.970671, 1.570796, 1.706749],accel_mss,speed_ms,0,blend_radius_m)
  movel([0.135606, -0.994795, -2.746567, -0.971027, 1.570796, 1.706403],accel_mss,speed_ms,0,blend_radius_m)
  movel([0.135231, -0.994840, -2.746554, -0.970995, 1.570796, 1.706027],accel_mss,speed_ms,0,blend_radius_m)
  movel([0.134795, -0.995087, -2.746482, -0.970820, 1.570796, 1.705592],accel_mss,speed_ms,0,blend_radius_m)
  movel([0.133917, -0.995925, -2.746236, -0.970228, 1.570796, 1.704713],accel_mss,speed_ms,0,blend_radius_m)
  movel([0.132686, -0.997519, -2.745768, -0.969102, 1.570796, 1.703482],accel_mss,speed_ms,0,blend_radius_m)
  movel([0.131708, -0.999114, -2.745297, -0.967978, 1.570796, 1.702505],accel_mss,speed_ms,0,blend_radius_m)
  movel([0.130937, -1.000704, -2.744826, -0.966859, 1.570796, 1.701733],accel_mss,speed_ms,0,blend_radius_m)
  movel([0.130326, -1.002283, -2.744356, -0.965750, 1.570796, 1.701122],accel_mss,speed_ms,0,blend_radius_m)
  movel([0.128511, -1.008508, -2.742485, -0.961395, 1.570796, 1.699307],accel_mss,speed_ms,0,blend_radius_m)
  movel([0.127266, -1.012186, -2.741366, -0.958837, 1.570796, 1.698062],accel_mss,speed_ms,0,blend_radius_m)
  movel([0.125795, -1.015892, -2.740228, -0.956269, 1.570796, 1.696591],accel_mss,speed_ms,0,blend_radius_m)
  movel([0.124038, -1.019608, -2.739076, -0.953705, 1.570796, 1.694835],accel_mss,speed_ms,0,blend_radius_m)
  movel([0.121941, -1.023302, -2.737920, -0.951167, 1.570796, 1.692737],accel_mss,speed_ms,0,blend_radius_m)
  movel([0.122563, -1.020546, -2.738783, -0.953060, 1.570796, 1.693359],accel_mss,speed_ms,0,blend_radius_m)
  movel([0.122553, -1.018087, -2.739548, -0.954753, 1.570796, 1.693350],accel_mss,speed_ms,0,blend_radius_m)
  movel([0.122409, -1.017556, -2.739713, -0.955120, 1.570796, 1.693205],accel_mss,speed_ms,0,blend_radius_m)
  movel([0.122040, -1.017264, -2.739804, -0.955321, 1.570796, 1.692837],accel_mss,speed_ms,0,blend_radius_m)
  movel([0.121554, -1.017348, -2.739778, -0.955263, 1.570796, 1.692350],accel_mss,speed_ms,0,blend_radius_m)
  movel([0.121001, -1.017681, -2.739675, -0.955034, 1.570796, 1.691797],accel_mss,speed_ms,0,blend_radius_m)
  movel([0.119921, -1.018735, -2.739347, -0.954307, 1.570796, 1.690717],accel_mss,speed_ms,0,blend_radius_m)
  movel([0.118765, -1.020249, -2.738876, -0.953264, 1.570796, 1.689561],accel_mss,speed_ms,0,blend_radius_m)
  movel([0.117777, -1.021824, -2.738384, -0.952181, 1.570796, 1.688573],accel_mss,speed_ms,0,blend_radius_m)
  movel([0.116176, -1.025060, -2.737366, -0.949963, 1.570796, 1.686972],accel_mss,speed_ms,0,blend_radius_m)
  movel([0.113543, -1.031437, -2.735336, -0.945616, 1.570796, 1.684339],accel_mss,speed_ms,0,blend_radius_m)
  movel([0.111823, -1.034987, -2.734192, -0.943210, 1.570796, 1.682619],accel_mss,speed_ms,0,blend_radius_m)
  movel([0.109889, -1.038516, -2.733044, -0.940829, 1.570796, 1.680686],accel_mss,speed_ms,0,blend_radius_m)
  movel([0.107694, -1.041973, -2.731910, -0.938505, 1.570796, 1.678490],accel_mss,speed_ms,0,blend_radius_m)
  movel([0.105191, -1.045314, -2.730805, -0.936269, 1.570796, 1.675988],accel_mss,speed_ms,0,blend_radius_m)
  movel([0.105698, -1.043796, -2.731309, -0.937284, 1.570796, 1.676494],accel_mss,speed_ms,0,blend_radius_m)
  movel([0.106188, -1.040939, -2.732251, -0.939199, 1.570796, 1.676984],accel_mss,speed_ms,0,blend_radius_m)
  movel([0.106161, -1.039642, -2.732676, -0.940071, 1.570796, 1.676958],accel_mss,speed_ms,0,blend_radius_m)
  movel([0.106006, -1.039134, -2.732842, -0.940413, 1.570796, 1.676802],accel_mss,speed_ms,0,blend_radius_m)
  movel([0.105552, -1.039029, -2.732877, -0.940483, 1.570796, 1.676348],accel_mss,speed_ms,0,blend_radius_m)
  movel([0.104890, -1.039542, -2.732709, -0.940138, 1.570796, 1.675687],accel_mss,speed_ms,0,blend_radius_m)
  movel([0.103405, -1.041178, -2.732172, -0.939039, 1.570796, 1.674202],accel_mss,speed_ms,0,blend_radius_m)
  movel([0.102119, -1.042843, -2.731623, -0.937922, 1.570796, 1.672915],accel_mss,speed_ms,0,blend_radius_m)
  movel([0.099909, -1.046239, -2.730498, -0.935652, 1.570796, 1.670705],accel_mss,speed_ms,0,blend_radius_m)
  movel([0.097790, -1.049665, -2.729352, -0.933372, 1.570796, 1.668586],accel_mss,speed_ms,0,blend_radius_m)
  movel([0.096618, -1.051374, -2.728777, -0.932238, 1.570796, 1.667414],accel_mss,speed_ms,0,blend_radius_m)
  movel([0.095292, -1.053072, -2.728204, -0.931113, 1.570796, 1.666088],accel_mss,speed_ms,0,blend_radius_m)
  movel([0.091838, -1.057004, -2.726866, -0.928519, 1.570796, 1.662635],accel_mss,speed_ms,0,blend_radius_m)
  movel([0.088265, -1.060789, -2.725566, -0.926034, 1.570796, 1.659061],accel_mss,speed_ms,0,blend_radius_m)
  movel([0.084609, -1.064431, -2.724303, -0.923654, 1.570796, 1.655405],accel_mss,speed_ms,0,blend_radius_m)
  movel([0.080897, -1.067952, -2.723072, -0.921365, 1.570796, 1.651693],accel_mss,speed_ms,0,blend_radius_m)
  speed_ms = 0.005
  movel([0.080897, -1.058391, -2.717670, -0.936328, 1.570796, 1.651693],accel_mss,speed_ms,0,blend_radius_m)
  speed_ms = 0.040
  movel([0.052585, -1.030085, -2.727167, -0.955137, 1.570796, 1.623381],accel_mss,speed_ms,0,blend_radius_m)
  speed_ms = 0.005
  movel([0.052585, -1.039609, -2.732687, -0.940093, 1.570796, 1.623381],accel_mss,speed_ms,0,blend_radius_m)
  speed_ms = 0.025
  movel([0.053739, -1.038256, -2.733129, -0.941004, 1.570796, 1.624535],accel_mss,speed_ms,0,blend_radius_m)
  movel([0.054770, -1.036784, -2.733609, -0.941996, 1.570796, 1.625566],accel_mss,speed_ms,0,blend_radius_m)
  movel([0.056627, -1.033615, -2.734635, -0.944139, 1.570796, 1.627423],accel_mss,speed_ms,0,blend_radius_m)
  movel([0.058462, -1.030371, -2.735678, -0.946341, 1.570796, 1.629259],accel_mss,speed_ms,0,blend_radius_m)
  movel([0.059472, -1.028801, -2.736179, -0.947409, 1.570796, 1.630269],accel_mss,speed_ms,0,blend_radius_m)
  movel([0.060595, -1.027315, -2.736652, -0.948422, 1.570796, 1.631391],accel_mss,speed_ms,0,blend_radius_m)
  movel([0.061493, -1.026328, -2.736965, -0.949096, 1.570796, 1.632289],accel_mss,speed_ms,0,blend_radius_m)
  movel([0.062238, -1.025695, -2.737165, -0.949529, 1.570796, 1.633034],accel_mss,speed_ms,0,blend_radius_m)
  movel([0.062844, -1.025377, -2.737266, -0.949747, 1.570796, 1.633640],accel_mss,speed_ms,0,blend_radius_m)
  movel([0.063327, -1.025333, -2.737279, -0.949776, 1.570796, 1.634123],accel_mss,speed_ms,0,blend_radius_m)
  movel([0.063959, -1.025948, -2.737085, -0.949356, 1.570796, 1.634756],accel_mss,speed_ms,0,blend_radius_m)
  movel([0.064238, -1.027239, -2.736676, -0.948474, 1.570796, 1.635035],accel_mss,speed_ms,0,blend_radius_m)
  movel([0.064127, -1.030691, -2.735575, -0.946123, 1.570796, 1.634924],accel_mss,speed_ms,0,blend_radius_m)
  movel([0.063808, -1.033367, -2.734715, -0.944307, 1.570796, 1.634605],accel_mss,speed_ms,0,blend_radius_m)
  movel([0.065855, -1.030129, -2.735755, -0.946505, 1.570796, 1.636651],accel_mss,speed_ms,0,blend_radius_m)
  movel([0.067407, -1.027030, -2.736742, -0.948617, 1.570796, 1.638203],accel_mss,speed_ms,0,blend_radius_m)
  movel([0.068592, -1.024022, -2.737693, -0.950674, 1.570796, 1.639389],accel_mss,speed_ms,0,blend_radius_m)
  movel([0.069527, -1.021071, -2.738619, -0.952699, 1.570796, 1.640323],accel_mss,speed_ms,0,blend_radius_m)
  movel([0.072078, -1.012124, -2.741385, -0.958880, 1.570796, 1.642875],accel_mss,speed_ms,0,blend_radius_m)
  movel([0.073262, -1.008964, -2.742347, -0.961078, 1.570796, 1.644059],accel_mss,speed_ms,0,blend_radius_m)
  movel([0.073925, -1.007674, -2.742738, -0.961977, 1.570796, 1.644722],accel_mss,speed_ms,0,blend_radius_m)
  movel([0.074609, -1.006839, -2.742990, -0.962560, 1.570796, 1.645405],accel_mss,speed_ms,0,blend_radius_m)
  movel([0.075288, -1.006394, -2.743124, -0.962871, 1.570796, 1.646084],accel_mss,speed_ms,0,blend_radius_m)
  movel([0.075933, -1.006282, -2.743158, -0.962949, 1.570796, 1.646729],accel_mss,speed_ms,0,blend_radius_m)
  movel([0.076523, -1.006435, -2.743111, -0.962842, 1.570796, 1.647320],accel_mss,speed_ms,0,blend_radius_m)
  movel([0.077028, -1.006794, -2.743003, -0.962592, 1.570796, 1.647824],accel_mss,speed_ms,0,blend_radius_m)
  movel([0.077688, -1.007869, -2.742679, -0.961841, 1.570796, 1.648484],accel_mss,speed_ms,0,blend_radius_m)
  movel([0.077828, -1.009308, -2.742243, -0.960839, 1.570796, 1.648624],accel_mss,speed_ms,0,blend_radius_m)
  movel([0.077674, -1.011309, -2.741634, -0.959446, 1.570796, 1.648471],accel_mss,speed_ms,0,blend_radius_m)
  movel([0.077147, -1.015098, -2.740473, -0.956819, 1.570796, 1.647943],accel_mss,speed_ms,0,blend_radius_m)
  movel([0.079247, -1.008913, -2.742363, -0.961113, 1.570796, 1.650044],accel_mss,speed_ms,0,blend_radius_m)
  movel([0.080045, -1.005879, -2.743279, -0.963231, 1.570796, 1.650842],accel_mss,speed_ms,0,blend_radius_m)
  movel([0.081117, -0.999980, -2.745041, -0.967368, 1.570796, 1.651913],accel_mss,speed_ms,0,blend_radius_m)
  movel([0.081382, -0.997146, -2.745878, -0.969366, 1.570796, 1.652178],accel_mss,speed_ms,0,blend_radius_m)
  movel([0.081355, -0.991769, -2.747449, -0.973171, 1.570796, 1.652151],accel_mss,speed_ms,0,blend_radius_m)
  speed_ms = 0.005
  movel([0.081355, -0.982372, -2.741737, -0.988280, 1.570796, 1.652151],accel_mss,speed_ms,0,blend_radius_m)
  speed_ms = 0.040
  movel([0.062258, -1.008565, -2.733955, -0.969869, 1.570796, 1.633054],accel_mss,speed_ms,0,blend_radius_m)
  speed_ms = 0.005
  movel([0.062258, -1.018041, -2.739563, -0.954785, 1.570796, 1.633054],accel_mss,speed_ms,0,blend_radius_m)
  speed_ms = 0.025
  movel([0.059858, -1.021752, -2.738406, -0.952231, 1.570796, 1.630654],accel_mss,speed_ms,0,blend_radius_m)
  movel([0.057669, -1.025486, -2.737231, -0.949671, 1.570796, 1.628466],accel_mss,speed_ms,0,blend_radius_m)
  movel([0.053440, -1.032916, -2.734861, -0.944613, 1.570796, 1.624237],accel_mss,speed_ms,0,blend_radius_m)
  movel([0.051127, -1.036589, -2.733672, -0.942128, 1.570796, 1.621923],accel_mss,speed_ms,0,blend_radius_m)
  movel([0.048566, -1.040150, -2.732510, -0.939730, 1.570796, 1.619362],accel_mss,speed_ms,0,blend_radius_m)
  movel([0.045728, -1.043458, -2.731420, -0.937511, 1.570796, 1.616525],accel_mss,speed_ms,0,blend_radius_m)
  movel([0.044200, -1.044973, -2.730919, -0.936498, 1.570796, 1.614997],accel_mss,speed_ms,0,blend_radius_m)
  movel([0.042596, -1.046373, -2.730453, -0.935563, 1.570796, 1.613392],accel_mss,speed_ms,0,blend_radius_m)
  movel([0.043768, -1.045118, -2.730870, -0.936401, 1.570796, 1.614565],accel_mss,speed_ms,0,blend_radius_m)
  movel([0.044992, -1.043309, -2.731470, -0.937610, 1.570796, 1.615788],accel_mss,speed_ms,0,blend_radius_m)
  movel([0.046127, -1.041201, -2.732165, -0.939024, 1.570796, 1.616923],accel_mss,speed_ms,0,blend_radius_m)
  movel([0.047012, -1.039061, -2.732866, -0.940462, 1.570796, 1.617809],accel_mss,speed_ms,0,blend_radius_m)
  movel([0.047502, -1.037150, -2.733490, -0.941750, 1.570796, 1.618298],accel_mss,speed_ms,0,blend_radius_m)
  movel([0.047545, -1.036370, -2.733743, -0.942276, 1.570796, 1.618341],accel_mss,speed_ms,0,blend_radius_m)
  movel([0.047433, -1.035747, -2.733946, -0.942697, 1.570796, 1.618230],accel_mss,speed_ms,0,blend_radius_m)
  movel([0.047146, -1.035314, -2.734086, -0.942989, 1.570796, 1.617942],accel_mss,speed_ms,0,blend_radius_m)
  movel([0.046658, -1.035113, -2.734151, -0.943125, 1.570796, 1.617455],accel_mss,speed_ms,0,blend_radius_m)
  movel([0.045960, -1.035169, -2.734133, -0.943087, 1.570796, 1.616756],accel_mss,speed_ms,0,blend_radius_m)
  movel([0.045023, -1.035521, -2.734019, -0.942849, 1.570796, 1.615819],accel_mss,speed_ms,0,blend_radius_m)
  movel([0.043517, -1.036548, -2.733685, -0.942156, 1.570796, 1.614313],accel_mss,speed_ms,0,blend_radius_m)
  movel([0.037327, -1.042105, -2.731867, -0.938417, 1.570796, 1.608124],accel_mss,speed_ms,0,blend_radius_m)
  movel([0.034681, -1.044212, -2.731171, -0.937006, 1.570796, 1.605478],accel_mss,speed_ms,0,blend_radius_m)
  movel([0.031966, -1.046152, -2.730527, -0.935710, 1.570796, 1.602762],accel_mss,speed_ms,0,blend_radius_m)
  movel([0.029266, -1.047819, -2.729971, -0.934599, 1.570796, 1.600063],accel_mss,speed_ms,0,blend_radius_m)
  movel([0.026666, -1.049095, -2.729544, -0.933751, 1.570796, 1.597462],accel_mss,speed_ms,0,blend_radius_m)
  movel([0.024244, -1.049870, -2.729283, -0.933235, 1.570796, 1.595040],accel_mss,speed_ms,0,blend_radius_m)
  movel([0.022086, -1.050024, -2.729232, -0.933133, 1.570796, 1.592882],accel_mss,speed_ms,0,blend_radius_m)
  movel([0.022777, -1.049867, -2.729284, -0.933237, 1.570796, 1.593573],accel_mss,speed_ms,0,blend_radius_m)
  movel([0.023686, -1.049351, -2.729458, -0.933580, 1.570796, 1.594482],accel_mss,speed_ms,0,blend_radius_m)
  movel([0.025867, -1.047613, -2.730040, -0.934737, 1.570796, 1.596664],accel_mss,speed_ms,0,blend_radius_m)
  movel([0.028010, -1.045547, -2.730728, -0.936114, 1.570796, 1.598806],accel_mss,speed_ms,0,blend_radius_m)
  movel([0.029486, -1.043905, -2.731273, -0.937212, 1.570796, 1.600282],accel_mss,speed_ms,0,blend_radius_m)
  movel([0.030353, -1.042650, -2.731687, -0.938052, 1.570796, 1.601149],accel_mss,speed_ms,0,blend_radius_m)
  movel([0.030677, -1.041821, -2.731960, -0.938607, 1.570796, 1.601473],accel_mss,speed_ms,0,blend_radius_m)
  movel([0.030544, -1.041351, -2.732115, -0.938923, 1.570796, 1.601341],accel_mss,speed_ms,0,blend_radius_m)
  movel([0.030055, -1.041173, -2.732174, -0.939042, 1.570796, 1.600851],accel_mss,speed_ms,0,blend_radius_m)
  movel([0.028394, -1.041421, -2.732092, -0.938876, 1.570796, 1.599190],accel_mss,speed_ms,0,blend_radius_m)
  movel([0.026468, -1.042023, -2.731894, -0.938472, 1.570796, 1.597264],accel_mss,speed_ms,0,blend_radius_m)
  movel([0.022092, -1.043388, -2.731444, -0.937558, 1.570796, 1.592888],accel_mss,speed_ms,0,blend_radius_m)
  movel([0.017739, -1.044375, -2.731117, -0.936897, 1.570796, 1.588535],accel_mss,speed_ms,0,blend_radius_m)
  movel([0.015686, -1.044593, -2.731045, -0.936751, 1.570796, 1.586482],accel_mss,speed_ms,0,blend_radius_m)
  movel([0.013777, -1.044552, -2.731058, -0.936779, 1.570796, 1.584574],accel_mss,speed_ms,0,blend_radius_m)
  movel([0.012060, -1.044196, -2.731176, -0.937017, 1.570796, 1.582856],accel_mss,speed_ms,0,blend_radius_m)
  movel([0.010581, -1.043471, -2.731416, -0.937502, 1.570796, 1.581377],accel_mss,speed_ms,0,blend_radius_m)
  movel([0.013190, -1.042629, -2.731694, -0.938066, 1.570796, 1.583987],accel_mss,speed_ms,0,blend_radius_m)
  movel([0.014621, -1.041860, -2.731948, -0.938582, 1.570796, 1.585417],accel_mss,speed_ms,0,blend_radius_m)
  movel([0.015257, -1.041357, -2.732113, -0.938919, 1.570796, 1.586053],accel_mss,speed_ms,0,blend_radius_m)
  movel([0.015800, -1.040757, -2.732310, -0.939322, 1.570796, 1.586596],accel_mss,speed_ms,0,blend_radius_m)
  movel([0.016023, -1.040300, -2.732460, -0.939629, 1.570796, 1.586820],accel_mss,speed_ms,0,blend_radius_m)
  movel([0.015994, -1.039885, -2.732596, -0.939907, 1.570796, 1.586790],accel_mss,speed_ms,0,blend_radius_m)
  movel([0.015315, -1.039176, -2.732828, -0.940384, 1.570796, 1.586112],accel_mss,speed_ms,0,blend_radius_m)
  movel([0.013996, -1.038617, -2.733011, -0.940761, 1.570796, 1.584792],accel_mss,speed_ms,0,blend_radius_m)
  movel([0.012280, -1.038185, -2.733152, -0.941052, 1.570796, 1.583076],accel_mss,speed_ms,0,blend_radius_m)
  movel([0.006259, -1.037325, -2.733433, -0.941631, 1.570796, 1.577055],accel_mss,speed_ms,0,blend_radius_m)
  movel([0.004079, -1.036662, -2.733648, -0.942079, 1.570796, 1.574875],accel_mss,speed_ms,0,blend_radius_m)
  movel([0.002111, -1.035693, -2.733963, -0.942733, 1.570796, 1.572908],accel_mss,speed_ms,0,blend_radius_m)
  movel([0.000486, -1.034331, -2.734404, -0.943654, 1.570796, 1.571283],accel_mss,speed_ms,0,blend_radius_m)
  movel([-0.000685, -1.032493, -2.734997, -0.944900, 1.570796, 1.570112],accel_mss,speed_ms,0,blend_radius_m)
  movel([0.001330, -1.033226, -2.734761, -0.944403, 1.570796, 1.572126],accel_mss,speed_ms,0,blend_radius_m)
  movel([0.002588, -1.033348, -2.734721, -0.944320, 1.570796, 1.573385],accel_mss,speed_ms,0,blend_radius_m)
  movel([0.003813, -1.033033, -2.734823, -0.944533, 1.570796, 1.574610],accel_mss,speed_ms,0,blend_radius_m)
  movel([0.004986, -1.032204, -2.735089, -0.945095, 1.570796, 1.575782],accel_mss,speed_ms,0,blend_radius_m)
  movel([0.005693, -1.031233, -2.735401, -0.945755, 1.570796, 1.576489],accel_mss,speed_ms,0,blend_radius_m)
  movel([0.005907, -1.030251, -2.735716, -0.946422, 1.570796, 1.576703],accel_mss,speed_ms,0,blend_radius_m)
  movel([0.005604, -1.029382, -2.735993, -0.947013, 1.570796, 1.576400],accel_mss,speed_ms,0,blend_radius_m)
  movel([0.003068, -1.025457, -2.737240, -0.949692, 1.570796, 1.573864],accel_mss,speed_ms,0,blend_radius_m)
  movel([0.001141, -1.021104, -2.738609, -0.952676, 1.570796, 1.571937],accel_mss,speed_ms,0,blend_radius_m)
  movel([0.000453, -1.018694, -2.739360, -0.954335, 1.570796, 1.571250],accel_mss,speed_ms,0,blend_radius_m)
  movel([-0.000030, -1.016091, -2.740166, -0.956132, 1.570796, 1.570766],accel_mss,speed_ms,0,blend_radius_m)
  movel([-0.000289, -1.013264, -2.741036, -0.958089, 1.570796, 1.570507],accel_mss,speed_ms,0,blend_radius_m)
  movel([-0.000305, -1.010182, -2.741977, -0.960230, 1.570796, 1.570491],accel_mss,speed_ms,0,blend_radius_m)
  speed_ms = 0.005
  movel([-0.000305, -1.000727, -2.736338, -0.975324, 1.570796, 1.570491],accel_mss,speed_ms,0,blend_radius_m)
  speed_ms = 0.040
  movel([-0.041269, -0.993146, -2.738598, -0.980645, 1.570796, 1.529527],accel_mss,speed_ms,0,blend_radius_m)
  speed_ms = 0.005
  movel([-0.041269, -1.002578, -2.744268, -0.965543, 1.570796, 1.529527],accel_mss,speed_ms,0,blend_radius_m)
  speed_ms = 0.025
  movel([-0.037935, -0.997017, -2.745915, -0.969456, 1.570796, 1.532862],accel_mss,speed_ms,0,blend_radius_m)
  movel([-0.034722, -0.991400, -2.747556, -0.973433, 1.570796, 1.536074],accel_mss,speed_ms,0,blend_radius_m)
  movel([-0.028597, -0.979963, -2.750824, -0.981601, 1.570796, 1.542199],accel_mss,speed_ms,0,blend_radius_m)
  movel([-0.022885, -0.968292, -2.754061, -0.990035, 1.570796, 1.547912],accel_mss,speed_ms,0,blend_radius_m)
  movel([-0.017602, -0.956425, -2.757254, -0.998710, 1.570796, 1.553194],accel_mss,speed_ms,0,blend_radius_m)
  movel([-0.012765, -0.944397, -2.760390, -1.007602, 1.570796, 1.558032],accel_mss,speed_ms,0,blend_radius_m)
  movel([-0.008393, -0.932256, -2.763456, -1.016677, 1.570796, 1.562403],accel_mss,speed_ms,0,blend_radius_m)
  movel([-0.004507, -0.920055, -2.766439, -1.025896, 1.570796, 1.566289],accel_mss,speed_ms,0,blend_radius_m)
  movel([-0.001128, -0.907838, -2.769328, -1.035222, 1.570796, 1.569668],accel_mss,speed_ms,0,blend_radius_m)
  movel([0.001717, -0.895676, -2.772111, -1.044602, 1.570796, 1.572514],accel_mss,speed_ms,0,blend_radius_m)
  movel([0.004003, -0.883627, -2.774778, -1.053984, 1.570796, 1.574800],accel_mss,speed_ms,0,blend_radius_m)
  movel([0.005699, -0.871763, -2.777318, -1.063308, 1.570796, 1.576495],accel_mss,speed_ms,0,blend_radius_m)
  movel([0.006772, -0.860158, -2.779722, -1.072509, 1.570796, 1.577568],accel_mss,speed_ms,0,blend_radius_m)
  movel([0.007201, -0.848881, -2.781983, -1.081525, 1.570796, 1.577998],accel_mss,speed_ms,0,blend_radius_m)
  movel([0.006944, -0.838026, -2.784091, -1.090272, 1.570796, 1.577741],accel_mss,speed_ms,0,blend_radius_m)
  movel([0.005975, -0.827674, -2.786040, -1.098675, 1.570796, 1.576771],accel_mss,speed_ms,0,blend_radius_m)
  movel([0.003369, -0.813036, -2.788697, -1.110657, 1.570796, 1.574166],accel_mss,speed_ms,0,blend_radius_m)
  movel([0.003313, -0.810302, -2.789180, -1.112908, 1.570796, 1.574110],accel_mss,speed_ms,0,blend_radius_m)
  movel([0.003753, -0.807229, -2.789718, -1.115442, 1.570796, 1.574550],accel_mss,speed_ms,0,blend_radius_m)
  movel([0.005074, -0.802618, -2.790517, -1.119254, 1.570796, 1.575870],accel_mss,speed_ms,0,blend_radius_m)
  movel([0.006722, -0.798785, -2.791173, -1.122432, 1.570796, 1.577519],accel_mss,speed_ms,0,blend_radius_m)
  movel([0.007652, -0.797149, -2.791450, -1.123790, 1.570796, 1.578448],accel_mss,speed_ms,0,blend_radius_m)
  movel([0.009696, -0.794389, -2.791915, -1.126085, 1.570796, 1.580493],accel_mss,speed_ms,0,blend_radius_m)
  movel([0.010791, -0.793265, -2.792103, -1.127021, 1.570796, 1.581587],accel_mss,speed_ms,0,blend_radius_m)
  movel([0.013113, -0.791473, -2.792402, -1.128514, 1.570796, 1.583910],accel_mss,speed_ms,0,blend_radius_m)
  movel([0.015556, -0.790256, -2.792604, -1.129529, 1.570796, 1.586352],accel_mss,speed_ms,0,blend_radius_m)
  movel([0.018066, -0.789559, -2.792719, -1.130111, 1.570796, 1.588863],accel_mss,speed_ms,0,blend_radius_m)
  movel([0.020598, -0.789326, -2.792757, -1.130306, 1.570796, 1.591395],accel_mss,speed_ms,0,blend_radius_m)
  movel([0.023097, -0.789495, -2.792729, -1.130165, 1.570796, 1.593894],accel_mss,speed_ms,0,blend_radius_m)
  movel([0.025518, -0.790012, -2.792644, -1.129733, 1.570796, 1.596315],accel_mss,speed_ms,0,blend_radius_m)
  movel([0.029924, -0.791821, -2.792344, -1.128224, 1.570796, 1.600720],accel_mss,speed_ms,0,blend_radius_m)
  movel([0.033447, -0.794254, -2.791937, -1.126198, 1.570796, 1.604244],accel_mss,speed_ms,0,blend_radius_m)
  movel([0.035752, -0.796766, -2.791515, -1.124108, 1.570796, 1.606548],accel_mss,speed_ms,0,blend_radius_m)
  movel([0.037774, -0.800397, -2.790898, -1.121094, 1.570796, 1.608570],accel_mss,speed_ms,0,blend_radius_m)
  movel([0.039406, -0.804424, -2.790206, -1.117760, 1.570796, 1.610203],accel_mss,speed_ms,0,blend_radius_m)
  movel([0.041880, -0.813222, -2.788663, -1.110503, 1.570796, 1.612676],accel_mss,speed_ms,0,blend_radius_m)
  movel([0.043907, -0.822340, -2.787022, -1.103027, 1.570796, 1.614703],accel_mss,speed_ms,0,blend_radius_m)
  movel([0.046189, -0.831001, -2.785420, -1.095967, 1.570796, 1.616985],accel_mss,speed_ms,0,blend_radius_m)
  movel([0.048787, -0.838196, -2.784059, -1.090135, 1.570796, 1.619584],accel_mss,speed_ms,0,blend_radius_m)
  movel([0.050495, -0.841348, -2.783453, -1.087588, 1.570796, 1.621292],accel_mss,speed_ms,0,blend_radius_m)
  movel([0.052701, -0.843939, -2.782951, -1.085499, 1.570796, 1.623497],accel_mss,speed_ms,0,blend_radius_m)
  movel([0.054025, -0.844791, -2.782785, -1.084813, 1.570796, 1.624822],accel_mss,speed_ms,0,blend_radius_m)
  movel([0.054860, -0.844951, -2.782754, -1.084684, 1.570796, 1.625656],accel_mss,speed_ms,0,blend_radius_m)
  movel([0.055847, -0.844825, -2.782779, -1.084786, 1.570796, 1.626643],accel_mss,speed_ms,0,blend_radius_m)
  movel([0.057282, -0.844187, -2.782903, -1.085299, 1.570796, 1.628078],accel_mss,speed_ms,0,blend_radius_m)
  movel([0.058791, -0.843135, -2.783107, -1.086147, 1.570796, 1.629587],accel_mss,speed_ms,0,blend_radius_m)
  movel([0.061813, -0.840324, -2.783650, -1.088415, 1.570796, 1.632609],accel_mss,speed_ms,0,blend_radius_m)
  movel([0.065119, -0.836744, -2.784336, -1.091310, 1.570796, 1.635915],accel_mss,speed_ms,0,blend_radius_m)
  movel([0.068277, -0.833009, -2.785043, -1.094337, 1.570796, 1.639073],accel_mss,speed_ms,0,blend_radius_m)
  movel([0.074274, -0.825176, -2.786502, -1.100711, 1.570796, 1.645070],accel_mss,speed_ms,0,blend_radius_m)
  movel([0.085956, -0.808860, -2.789433, -1.114096, 1.570796, 1.656752],accel_mss,speed_ms,0,blend_radius_m)
  movel([0.091724, -0.801228, -2.790756, -1.120405, 1.570796, 1.662520],accel_mss,speed_ms,0,blend_radius_m)
  movel([0.095118, -0.797086, -2.791461, -1.123842, 1.570796, 1.665914],accel_mss,speed_ms,0,blend_radius_m)
  movel([0.098550, -0.793336, -2.792091, -1.126962, 1.570796, 1.669346],accel_mss,speed_ms,0,blend_radius_m)
  movel([0.100208, -0.791749, -2.792356, -1.128284, 1.570796, 1.671005],accel_mss,speed_ms,0,blend_radius_m)
  movel([0.101792, -0.790433, -2.792574, -1.129382, 1.570796, 1.672589],accel_mss,speed_ms,0,blend_radius_m)
  movel([0.103267, -0.789446, -2.792738, -1.130206, 1.570796, 1.674063],accel_mss,speed_ms,0,blend_radius_m)
  movel([0.104605, -0.788849, -2.792836, -1.130704, 1.570796, 1.675402],accel_mss,speed_ms,0,blend_radius_m)
  movel([0.105774, -0.788696, -2.792861, -1.130832, 1.570796, 1.676571],accel_mss,speed_ms,0,blend_radius_m)
  movel([0.106748, -0.789041, -2.792804, -1.130543, 1.570796, 1.677544],accel_mss,speed_ms,0,blend_radius_m)
  movel([0.107496, -0.789949, -2.792654, -1.129786, 1.570796, 1.678292],accel_mss,speed_ms,0,blend_radius_m)
  movel([0.107985, -0.791473, -2.792402, -1.128514, 1.570796, 1.678781],accel_mss,speed_ms,0,blend_radius_m)
  movel([0.108380, -0.794563, -2.791886, -1.125941, 1.570796, 1.679177],accel_mss,speed_ms,0,blend_radius_m)
  movel([0.108432, -0.797834, -2.791334, -1.123221, 1.570796, 1.679228],accel_mss,speed_ms,0,blend_radius_m)
  movel([0.108163, -0.801260, -2.790750, -1.120379, 1.570796, 1.678960],accel_mss,speed_ms,0,blend_radius_m)
  movel([0.107597, -0.804831, -2.790135, -1.117423, 1.570796, 1.678393],accel_mss,speed_ms,0,blend_radius_m)
  movel([0.106747, -0.808517, -2.789493, -1.114379, 1.570796, 1.677543],accel_mss,speed_ms,0,blend_radius_m)
  movel([0.105636, -0.812303, -2.788826, -1.111259, 1.570796, 1.676432],accel_mss,speed_ms,0,blend_radius_m)
  movel([0.104281, -0.816174, -2.788137, -1.108078, 1.570796, 1.675078],accel_mss,speed_ms,0,blend_radius_m)
  movel([0.102705, -0.820110, -2.787427, -1.104851, 1.570796, 1.673502],accel_mss,speed_ms,0,blend_radius_m)
  movel([0.098963, -0.828104, -2.785961, -1.098325, 1.570796, 1.669759],accel_mss,speed_ms,0,blend_radius_m)
  movel([0.094548, -0.836162, -2.784446, -1.091780, 1.570796, 1.665345],accel_mss,speed_ms,0,blend_radius_m)
  movel([0.089597, -0.844162, -2.782908, -1.085319, 1.570796, 1.660394],accel_mss,speed_ms,0,blend_radius_m)
  movel([0.084252, -0.851984, -2.781368, -1.079037, 1.570796, 1.655048],accel_mss,speed_ms,0,blend_radius_m)
  movel([0.071998, -0.869001, -2.777898, -1.065490, 1.570796, 1.642794],accel_mss,speed_ms,0,blend_radius_m)
  movel([0.065571, -0.877247, -2.776155, -1.058987, 1.570796, 1.636367],accel_mss,speed_ms,0,blend_radius_m)
  movel([0.062299, -0.881107, -2.775325, -1.055957, 1.570796, 1.633095],accel_mss,speed_ms,0,blend_radius_m)
  movel([0.058990, -0.884724, -2.774539, -1.053126, 1.570796, 1.629786],accel_mss,speed_ms,0,blend_radius_m)
  movel([0.056838, -0.886874, -2.774068, -1.051447, 1.570796, 1.627635],accel_mss,speed_ms,0,blend_radius_m)
  movel([0.054684, -0.888815, -2.773641, -1.049933, 1.570796, 1.625481],accel_mss,speed_ms,0,blend_radius_m)
  movel([0.052541, -0.890518, -2.773264, -1.048607, 1.570796, 1.623337],accel_mss,speed_ms,0,blend_radius_m)
  movel([0.050425, -0.891949, -2.772946, -1.047494, 1.570796, 1.621221],accel_mss,speed_ms,0,blend_radius_m)
  movel([0.048357, -0.893077, -2.772694, -1.046618, 1.570796, 1.619154],accel_mss,speed_ms,0,blend_radius_m)
  movel([0.046350, -0.893870, -2.772517, -1.046002, 1.570796, 1.617147],accel_mss,speed_ms,0,blend_radius_m)
  movel([0.044425, -0.894289, -2.772423, -1.045677, 1.570796, 1.615221],accel_mss,speed_ms,0,blend_radius_m)
  movel([0.042592, -0.894302, -2.772420, -1.045667, 1.570796, 1.613389],accel_mss,speed_ms,0,blend_radius_m)
  movel([0.040937, -0.893875, -2.772516, -1.045998, 1.570796, 1.611733],accel_mss,speed_ms,0,blend_radius_m)
  movel([0.039563, -0.893092, -2.772691, -1.046606, 1.570796, 1.610360],accel_mss,speed_ms,0,blend_radius_m)
  movel([0.034961, -0.888743, -2.773657, -1.049989, 1.570796, 1.605758],accel_mss,speed_ms,0,blend_radius_m)
  movel([0.033548, -0.887950, -2.773832, -1.050607, 1.570796, 1.604344],accel_mss,speed_ms,0,blend_radius_m)
  movel([0.031832, -0.887524, -2.773926, -1.050940, 1.570796, 1.602629],accel_mss,speed_ms,0,blend_radius_m)
  movel([0.031048, -0.887630, -2.773902, -1.050857, 1.570796, 1.601844],accel_mss,speed_ms,0,blend_radius_m)
  movel([0.030681, -0.888132, -2.773792, -1.050466, 1.570796, 1.601477],accel_mss,speed_ms,0,blend_radius_m)
  movel([0.030199, -0.889279, -2.773538, -1.049571, 1.570796, 1.600996],accel_mss,speed_ms,0,blend_radius_m)
  movel([0.028942, -0.893177, -2.772672, -1.046540, 1.570796, 1.599739],accel_mss,speed_ms,0,blend_radius_m)
  movel([0.025811, -0.904798, -2.770033, -1.037558, 1.570796, 1.596608],accel_mss,speed_ms,0,blend_radius_m)
  movel([0.020960, -0.923948, -2.765497, -1.022943, 1.570796, 1.591756],accel_mss,speed_ms,0,blend_radius_m)
  movel([0.017470, -0.934196, -2.762973, -1.015220, 1.570796, 1.588266],accel_mss,speed_ms,0,blend_radius_m)
  movel([0.013608, -0.944412, -2.760386, -1.007591, 1.570796, 1.584404],accel_mss,speed_ms,0,blend_radius_m)
  movel([0.009426, -0.954566, -2.757745, -1.000078, 1.570796, 1.580223],accel_mss,speed_ms,0,blend_radius_m)
  movel([0.004989, -0.964618, -2.755060, -0.992710, 1.570796, 1.575785],accel_mss,speed_ms,0,blend_radius_m)
  movel([-0.000886, -0.977324, -2.751565, -0.983500, 1.570796, 1.569910],accel_mss,speed_ms,0,blend_radius_m)
  movel([-0.006924, -0.989870, -2.747999, -0.974520, 1.570796, 1.563873],accel_mss,speed_ms,0,blend_radius_m)
  movel([-0.013170, -1.002213, -2.744377, -0.965799, 1.570796, 1.557626],accel_mss,speed_ms,0,blend_radius_m)
  movel([-0.019682, -1.014308, -2.740716, -0.957365, 1.570796, 1.551114],accel_mss,speed_ms,0,blend_radius_m)
  movel([-0.026507, -1.026109, -2.737034, -0.949246, 1.570796, 1.544290],accel_mss,speed_ms,0,blend_radius_m)
  movel([-0.030048, -1.031887, -2.735191, -0.945311, 1.570796, 1.540749],accel_mss,speed_ms,0,blend_radius_m)
  movel([-0.033689, -1.037581, -2.733349, -0.941459, 1.570796, 1.537107],accel_mss,speed_ms,0,blend_radius_m)
  movel([-0.037435, -1.043186, -2.731510, -0.937693, 1.570796, 1.533362],accel_mss,speed_ms,0,blend_radius_m)
  movel([-0.041287, -1.048693, -2.729678, -0.934018, 1.570796, 1.529509],accel_mss,speed_ms,0,blend_radius_m)
  movel([-0.045255, -1.054106, -2.727853, -0.930430, 1.570796, 1.525541],accel_mss,speed_ms,0,blend_radius_m)
  movel([-0.049349, -1.059416, -2.726039, -0.926934, 1.570796, 1.521448],accel_mss,speed_ms,0,blend_radius_m)
  movel([-0.054352, -1.065585, -2.723901, -0.922903, 1.570796, 1.516444],accel_mss,speed_ms,0,blend_radius_m)
  movel([-0.056958, -1.068547, -2.722863, -0.920979, 1.570796, 1.513838],accel_mss,speed_ms,0,blend_radius_m)
  movel([-0.061649, -1.073305, -2.721180, -0.917904, 1.570796, 1.509147],accel_mss,speed_ms,0,blend_radius_m)
  movel([-0.064077, -1.075476, -2.720405, -0.916507, 1.570796, 1.506719],accel_mss,speed_ms,0,blend_radius_m)
  movel([-0.066519, -1.077212, -2.719783, -0.915394, 1.570796, 1.504277],accel_mss,speed_ms,0,blend_radius_m)
  movel([-0.067609, -1.077706, -2.719605, -0.915077, 1.570796, 1.503188],accel_mss,speed_ms,0,blend_radius_m)
  movel([-0.068545, -1.077845, -2.719556, -0.914989, 1.570796, 1.502251],accel_mss,speed_ms,0,blend_radius_m)
  movel([-0.067892, -1.075254, -2.720485, -0.916650, 1.570796, 1.502904],accel_mss,speed_ms,0,blend_radius_m)
  movel([-0.067596, -1.072798, -2.721360, -0.918231, 1.570796, 1.503200],accel_mss,speed_ms,0,blend_radius_m)
  movel([-0.067673, -1.071738, -2.721736, -0.918915, 1.570796, 1.503124],accel_mss,speed_ms,0,blend_radius_m)
  movel([-0.067948, -1.070854, -2.722049, -0.919486, 1.570796, 1.502849],accel_mss,speed_ms,0,blend_radius_m)
  movel([-0.068456, -1.070189, -2.722284, -0.919915, 1.570796, 1.502340],accel_mss,speed_ms,0,blend_radius_m)
  movel([-0.069242, -1.069801, -2.722421, -0.920166, 1.570796, 1.501554],accel_mss,speed_ms,0,blend_radius_m)
  movel([-0.071652, -1.069575, -2.722501, -0.920313, 1.570796, 1.499145],accel_mss,speed_ms,0,blend_radius_m)
  movel([-0.072322, -1.069232, -2.722622, -0.920535, 1.570796, 1.498475],accel_mss,speed_ms,0,blend_radius_m)
  movel([-0.072785, -1.068674, -2.722818, -0.920897, 1.570796, 1.498011],accel_mss,speed_ms,0,blend_radius_m)
  movel([-0.073179, -1.067056, -2.723387, -0.921947, 1.570796, 1.497617],accel_mss,speed_ms,0,blend_radius_m)
  movel([-0.073051, -1.065001, -2.724105, -0.923283, 1.570796, 1.497746],accel_mss,speed_ms,0,blend_radius_m)
  movel([-0.072608, -1.062800, -2.724870, -0.924719, 1.570796, 1.498188],accel_mss,speed_ms,0,blend_radius_m)
  movel([-0.070858, -1.056018, -2.727203, -0.929169, 1.570796, 1.499938],accel_mss,speed_ms,0,blend_radius_m)
  movel([-0.068698, -1.049004, -2.729574, -0.933811, 1.570796, 1.502098],accel_mss,speed_ms,0,blend_radius_m)
  movel([-0.067395, -1.045426, -2.730768, -0.936195, 1.570796, 1.503402],accel_mss,speed_ms,0,blend_radius_m)
  movel([-0.065910, -1.041806, -2.731965, -0.938617, 1.570796, 1.504886],accel_mss,speed_ms,0,blend_radius_m)
  movel([-0.064215, -1.038155, -2.733162, -0.941072, 1.570796, 1.506582],accel_mss,speed_ms,0,blend_radius_m)
  movel([-0.062279, -1.034474, -2.734358, -0.943558, 1.570796, 1.508517],accel_mss,speed_ms,0,blend_radius_m)
  movel([-0.060072, -1.030919, -2.735502, -0.945968, 1.570796, 1.510725],accel_mss,speed_ms,0,blend_radius_m)
  movel([-0.052653, -1.020644, -2.738753, -0.952992, 1.570796, 1.518143],accel_mss,speed_ms,0,blend_radius_m)
  movel([-0.046893, -1.011711, -2.741511, -0.959167, 1.570796, 1.523903],accel_mss,speed_ms,0,blend_radius_m)
  movel([-0.041269, -1.002578, -2.744268, -0.965543, 1.570796, 1.529527],accel_mss,speed_ms,0,blend_radius_m)
  movel([-0.038775, -0.998416, -2.745503, -0.968470, 1.570796, 1.532021],accel_mss,speed_ms,0,blend_radius_m)
  speed_ms = 0.005
  movel([-0.038775, -0.988997, -2.739817, -0.983575, 1.570796, 1.532021],accel_mss,speed_ms,0,blend_radius_m)
  speed_ms = 0.040
  movel([-0.089816, -1.062599, -2.716201, -0.933589, 1.570796, 1.480980],accel_mss,speed_ms,0,blend_radius_m)
  speed_ms = 0.005
  movel([-0.089816, -1.072164, -2.721585, -0.918639, 1.570796, 1.480980],accel_mss,speed_ms,0,blend_radius_m)
  speed_ms = 0.025
  movel([-0.085381, -1.075207, -2.720502, -0.916681, 1.570796, 1.485415],accel_mss,speed_ms,0,blend_radius_m)
  movel([-0.083192, -1.077028, -2.719849, -0.915512, 1.570796, 1.487604],accel_mss,speed_ms,0,blend_radius_m)
  movel([-0.081191, -1.079091, -2.719107, -0.914192, 1.570796, 1.489606],accel_mss,speed_ms,0,blend_radius_m)
  movel([-0.079489, -1.081409, -2.718268, -0.912712, 1.570796, 1.491307],accel_mss,speed_ms,0,blend_radius_m)
  movel([-0.078209, -1.084004, -2.717323, -0.911062, 1.570796, 1.492587],accel_mss,speed_ms,0,blend_radius_m)
  movel([-0.077467, -1.086898, -2.716262, -0.909229, 1.570796, 1.493329],accel_mss,speed_ms,0,blend_radius_m)
  movel([-0.077335, -1.088465, -2.715685, -0.908239, 1.570796, 1.493461],accel_mss,speed_ms,0,blend_radius_m)
  movel([-0.077380, -1.090110, -2.715076, -0.907203, 1.570796, 1.493416],accel_mss,speed_ms,0,blend_radius_m)
  movel([-0.078452, -1.089801, -2.715191, -0.907397, 1.570796, 1.492345],accel_mss,speed_ms,0,blend_radius_m)
  movel([-0.079150, -1.089214, -2.715408, -0.907767, 1.570796, 1.491646],accel_mss,speed_ms,0,blend_radius_m)
  movel([-0.080624, -1.087807, -2.715928, -0.908655, 1.570796, 1.490172],accel_mss,speed_ms,0,blend_radius_m)
  movel([-0.082650, -1.086807, -2.716296, -0.909286, 1.570796, 1.488147],accel_mss,speed_ms,0,blend_radius_m)
  movel([-0.084885, -1.086084, -2.716561, -0.909744, 1.570796, 1.485911],accel_mss,speed_ms,0,blend_radius_m)
  movel([-0.087305, -1.085624, -2.716730, -0.910035, 1.570796, 1.483491],accel_mss,speed_ms,0,blend_radius_m)
  movel([-0.089883, -1.085421, -2.716805, -0.910164, 1.570796, 1.480913],accel_mss,speed_ms,0,blend_radius_m)
  movel([-0.092594, -1.085463, -2.716789, -0.910137, 1.570796, 1.478203],accel_mss,speed_ms,0,blend_radius_m)
  movel([-0.095409, -1.085744, -2.716686, -0.909959, 1.570796, 1.475387],accel_mss,speed_ms,0,blend_radius_m)
  movel([-0.098307, -1.086257, -2.716498, -0.909634, 1.570796, 1.472490],accel_mss,speed_ms,0,blend_radius_m)
  movel([-0.101256, -1.086985, -2.716230, -0.909174, 1.570796, 1.469540],accel_mss,speed_ms,0,blend_radius_m)
  movel([-0.103243, -1.087638, -2.715990, -0.908761, 1.570796, 1.467553],accel_mss,speed_ms,0,blend_radius_m)
  movel([-0.104813, -1.088354, -2.715726, -0.908309, 1.570796, 1.465983],accel_mss,speed_ms,0,blend_radius_m)
  movel([-0.105996, -1.089120, -2.715443, -0.907826, 1.570796, 1.464800],accel_mss,speed_ms,0,blend_radius_m)
  movel([-0.106828, -1.089925, -2.715145, -0.907319, 1.570796, 1.463969],accel_mss,speed_ms,0,blend_radius_m)
  movel([-0.107346, -1.090767, -2.714833, -0.906789, 1.570796, 1.463451],accel_mss,speed_ms,0,blend_radius_m)
  movel([-0.107582, -1.091635, -2.714510, -0.906244, 1.570796, 1.463214],accel_mss,speed_ms,0,blend_radius_m)
  movel([-0.107579, -1.092525, -2.714178, -0.905685, 1.570796, 1.463218],accel_mss,speed_ms,0,blend_radius_m)
  movel([-0.107365, -1.093427, -2.713842, -0.905120, 1.570796, 1.463432],accel_mss,speed_ms,0,blend_radius_m)
  movel([-0.106462, -1.095245, -2.713161, -0.903983, 1.570796, 1.464334],accel_mss,speed_ms,0,blend_radius_m)
  movel([-0.102469, -1.100347, -2.711234, -0.900807, 1.570796, 1.468328],accel_mss,speed_ms,0,blend_radius_m)
  movel([-0.105068, -1.099441, -2.711578, -0.901369, 1.570796, 1.465728],accel_mss,speed_ms,0,blend_radius_m)
  movel([-0.110164, -1.097501, -2.712312, -0.902576, 1.570796, 1.460632],accel_mss,speed_ms,0,blend_radius_m)
  movel([-0.113027, -1.097016, -2.712495, -0.902878, 1.570796, 1.457770],accel_mss,speed_ms,0,blend_radius_m)
  movel([-0.116461, -1.096954, -2.712518, -0.902917, 1.570796, 1.454335],accel_mss,speed_ms,0,blend_radius_m)
  movel([-0.120018, -1.097104, -2.712462, -0.902823, 1.570796, 1.450778],accel_mss,speed_ms,0,blend_radius_m)
  movel([-0.127213, -1.097575, -2.712284, -0.902530, 1.570796, 1.443583],accel_mss,speed_ms,0,blend_radius_m)
  movel([-0.130713, -1.097667, -2.712250, -0.902473, 1.570796, 1.440083],accel_mss,speed_ms,0,blend_radius_m)
  movel([-0.134055, -1.097509, -2.712309, -0.902571, 1.570796, 1.436742],accel_mss,speed_ms,0,blend_radius_m)
  movel([-0.137170, -1.096991, -2.712504, -0.902893, 1.570796, 1.433626],accel_mss,speed_ms,0,blend_radius_m)
  movel([-0.139995, -1.095992, -2.712881, -0.903517, 1.570796, 1.430802],accel_mss,speed_ms,0,blend_radius_m)
  movel([-0.137192, -1.100505, -2.711174, -0.900709, 1.570796, 1.433605],accel_mss,speed_ms,0,blend_radius_m)
  movel([-0.135602, -1.102684, -2.710344, -0.899361, 1.570796, 1.435194],accel_mss,speed_ms,0,blend_radius_m)
  movel([-0.133826, -1.104407, -2.709685, -0.898298, 1.570796, 1.436971],accel_mss,speed_ms,0,blend_radius_m)
  movel([-0.136672, -1.103535, -2.710019, -0.898835, 1.570796, 1.434124],accel_mss,speed_ms,0,blend_radius_m)
  movel([-0.139763, -1.103035, -2.710210, -0.899144, 1.570796, 1.431033],accel_mss,speed_ms,0,blend_radius_m)
  movel([-0.146189, -1.102417, -2.710446, -0.899526, 1.570796, 1.424608],accel_mss,speed_ms,0,blend_radius_m)
  movel([-0.148233, -1.102031, -2.710593, -0.899764, 1.570796, 1.422563],accel_mss,speed_ms,0,blend_radius_m)
  movel([-0.150068, -1.101422, -2.710825, -0.900141, 1.570796, 1.420728],accel_mss,speed_ms,0,blend_radius_m)
  movel([-0.153333, -1.099751, -2.711461, -0.901177, 1.570796, 1.417463],accel_mss,speed_ms,0,blend_radius_m)
  movel([-0.156453, -1.097870, -2.712173, -0.902346, 1.570796, 1.414344],accel_mss,speed_ms,0,blend_radius_m)
  movel([-0.159894, -1.096258, -2.712780, -0.903350, 1.570796, 1.410903],accel_mss,speed_ms,0,blend_radius_m)
  movel([-0.161112, -1.095929, -2.712904, -0.903556, 1.570796, 1.409685],accel_mss,speed_ms,0,blend_radius_m)
  movel([-0.162467, -1.095832, -2.712941, -0.903616, 1.570796, 1.408329],accel_mss,speed_ms,0,blend_radius_m)
  movel([-0.163937, -1.096118, -2.712833, -0.903438, 1.570796, 1.406859],accel_mss,speed_ms,0,blend_radius_m)
  movel([-0.164701, -1.096444, -2.712710, -0.903235, 1.570796, 1.406095],accel_mss,speed_ms,0,blend_radius_m)
  movel([-0.165483, -1.096923, -2.712530, -0.902936, 1.570796, 1.405313],accel_mss,speed_ms,0,blend_radius_m)
  movel([-0.166307, -1.097594, -2.712277, -0.902518, 1.570796, 1.404490],accel_mss,speed_ms,0,blend_radius_m)
  movel([-0.167031, -1.098359, -2.711988, -0.902042, 1.570796, 1.403765],accel_mss,speed_ms,0,blend_radius_m)
  movel([-0.168230, -1.100097, -2.711330, -0.900963, 1.570796, 1.402566],accel_mss,speed_ms,0,blend_radius_m)
  movel([-0.169139, -1.101971, -2.710616, -0.899801, 1.570796, 1.401658],accel_mss,speed_ms,0,blend_radius_m)
  movel([-0.169815, -1.103820, -2.709909, -0.898659, 1.570796, 1.400982],accel_mss,speed_ms,0,blend_radius_m)
  movel([-0.170869, -1.101549, -2.710777, -0.900063, 1.570796, 1.399927],accel_mss,speed_ms,0,blend_radius_m)
  movel([-0.172146, -1.099518, -2.711549, -0.901322, 1.570796, 1.398650],accel_mss,speed_ms,0,blend_radius_m)
  movel([-0.175130, -1.095934, -2.712902, -0.903552, 1.570796, 1.395666],accel_mss,speed_ms,0,blend_radius_m)
  movel([-0.178288, -1.092531, -2.714176, -0.905682, 1.570796, 1.392508],accel_mss,speed_ms,0,blend_radius_m)
  movel([-0.181130, -1.088747, -2.715580, -0.908061, 1.570796, 1.389666],accel_mss,speed_ms,0,blend_radius_m)
  movel([-0.181947, -1.087017, -2.716218, -0.909153, 1.570796, 1.388849],accel_mss,speed_ms,0,blend_radius_m)
  movel([-0.182498, -1.085015, -2.716953, -0.910421, 1.570796, 1.388298],accel_mss,speed_ms,0,blend_radius_m)
  movel([-0.182819, -1.082793, -2.717765, -0.911832, 1.570796, 1.387977],accel_mss,speed_ms,0,blend_radius_m)
  movel([-0.182952, -1.080413, -2.718629, -0.913348, 1.570796, 1.387845],accel_mss,speed_ms,0,blend_radius_m)
  movel([-0.182776, -1.075380, -2.720440, -0.916570, 1.570796, 1.388020],accel_mss,speed_ms,0,blend_radius_m)
  movel([-0.182269, -1.070376, -2.722218, -0.919794, 1.570796, 1.388528],accel_mss,speed_ms,0,blend_radius_m)
  speed_ms = 0.005
  movel([-0.182269, -1.060813, -2.716826, -0.934750, 1.570796, 1.388528],accel_mss,speed_ms,0,blend_radius_m)
  speed_ms = 0.040
  # Splitting Linear movement in 2 (instruction 806: MoveL 765)
  movel([-0.154336, -0.986170, -2.740640, -0.985579, 1.570796, 1.416460],accel_mss,speed_ms,0,blend_radius_m)
  movel([-0.121695, -0.902275, -2.762511, -1.047602, 1.570796, 1.449101],accel_mss,speed_ms,0,blend_radius_m)
  speed_ms = 0.005
  movel([-0.121695, -0.911274, -2.768525, -1.032590, 1.570796, 1.449101],accel_mss,speed_ms,0,blend_radius_m)
  speed_ms = 0.025
  movel([-0.123729, -0.913790, -2.767933, -1.030667, 1.570796, 1.447067],accel_mss,speed_ms,0,blend_radius_m)
  movel([-0.123869, -0.914204, -2.767835, -1.030351, 1.570796, 1.446928],accel_mss,speed_ms,0,blend_radius_m)
  movel([-0.123677, -0.914661, -2.767726, -1.030002, 1.570796, 1.447119],accel_mss,speed_ms,0,blend_radius_m)
  movel([-0.122387, -0.915713, -2.767477, -1.029200, 1.570796, 1.448409],accel_mss,speed_ms,0,blend_radius_m)
  movel([-0.116786, -0.918278, -2.766865, -1.027246, 1.570796, 1.454011],accel_mss,speed_ms,0,blend_radius_m)
  movel([-0.108296, -0.921322, -2.766133, -1.024934, 1.570796, 1.462501],accel_mss,speed_ms,0,blend_radius_m)
  movel([-0.098262, -0.924654, -2.765326, -1.022410, 1.570796, 1.472535],accel_mss,speed_ms,0,blend_radius_m)
  movel([-0.078691, -0.931099, -2.763743, -1.017547, 1.570796, 1.492105],accel_mss,speed_ms,0,blend_radius_m)
  movel([-0.067694, -0.934660, -2.762857, -1.014872, 1.570796, 1.503103],accel_mss,speed_ms,0,blend_radius_m)
  movel([-0.066628, -0.934828, -2.762815, -1.014747, 1.570796, 1.504168],accel_mss,speed_ms,0,blend_radius_m)
  movel([-0.065426, -0.934741, -2.762836, -1.014811, 1.570796, 1.505370],accel_mss,speed_ms,0,blend_radius_m)
  movel([-0.064169, -0.934248, -2.762960, -1.015181, 1.570796, 1.506628],accel_mss,speed_ms,0,blend_radius_m)
  movel([-0.063539, -0.933804, -2.763070, -1.015514, 1.570796, 1.507257],accel_mss,speed_ms,0,blend_radius_m)
  movel([-0.062925, -0.933198, -2.763221, -1.015969, 1.570796, 1.507871],accel_mss,speed_ms,0,blend_radius_m)
  movel([-0.062039, -0.931894, -2.763546, -1.016949, 1.570796, 1.508758],accel_mss,speed_ms,0,blend_radius_m)
  movel([-0.061407, -0.930528, -2.763884, -1.017977, 1.570796, 1.509389],accel_mss,speed_ms,0,blend_radius_m)
  movel([-0.058516, -0.922949, -2.765740, -1.023700, 1.570796, 1.512280],accel_mss,speed_ms,0,blend_radius_m)
  movel([-0.056125, -0.915443, -2.767541, -1.029405, 1.570796, 1.514671],accel_mss,speed_ms,0,blend_radius_m)
  movel([-0.054216, -0.908045, -2.769280, -1.035063, 1.570796, 1.516580],accel_mss,speed_ms,0,blend_radius_m)
  movel([-0.052750, -0.900783, -2.770954, -1.040652, 1.570796, 1.518046],accel_mss,speed_ms,0,blend_radius_m)
  movel([-0.051705, -0.893685, -2.772558, -1.046145, 1.570796, 1.519091],accel_mss,speed_ms,0,blend_radius_m)
  movel([-0.051044, -0.886779, -2.774089, -1.051521, 1.570796, 1.519752],accel_mss,speed_ms,0,blend_radius_m)
  movel([-0.050737, -0.880094, -2.775544, -1.056752, 1.570796, 1.520059],accel_mss,speed_ms,0,blend_radius_m)
  movel([-0.050750, -0.873665, -2.776917, -1.061807, 1.570796, 1.520046],accel_mss,speed_ms,0,blend_radius_m)
  movel([-0.050960, -0.870879, -2.777504, -1.064006, 1.570796, 1.519836],accel_mss,speed_ms,0,blend_radius_m)
  movel([-0.051433, -0.868471, -2.778008, -1.065910, 1.570796, 1.519363],accel_mss,speed_ms,0,blend_radius_m)
  movel([-0.052166, -0.866437, -2.778431, -1.067521, 1.570796, 1.518631],accel_mss,speed_ms,0,blend_radius_m)
  movel([-0.053142, -0.864764, -2.778778, -1.068848, 1.570796, 1.517655],accel_mss,speed_ms,0,blend_radius_m)
  movel([-0.054358, -0.863451, -2.779048, -1.069890, 1.570796, 1.516439],accel_mss,speed_ms,0,blend_radius_m)
  movel([-0.055805, -0.862493, -2.779245, -1.070651, 1.570796, 1.514992],accel_mss,speed_ms,0,blend_radius_m)
  movel([-0.057470, -0.861872, -2.779372, -1.071145, 1.570796, 1.513326],accel_mss,speed_ms,0,blend_radius_m)
  movel([-0.059349, -0.861584, -2.779431, -1.071374, 1.570796, 1.511448],accel_mss,speed_ms,0,blend_radius_m)
  movel([-0.061426, -0.861621, -2.779423, -1.071345, 1.570796, 1.509370],accel_mss,speed_ms,0,blend_radius_m)
  movel([-0.063692, -0.861971, -2.779352, -1.071066, 1.570796, 1.507104],accel_mss,speed_ms,0,blend_radius_m)
  movel([-0.066142, -0.862623, -2.779218, -1.070548, 1.570796, 1.504655],accel_mss,speed_ms,0,blend_radius_m)
  movel([-0.068755, -0.863568, -2.779024, -1.069797, 1.570796, 1.502042],accel_mss,speed_ms,0,blend_radius_m)
  movel([-0.074446, -0.866290, -2.778462, -1.067637, 1.570796, 1.496350],accel_mss,speed_ms,0,blend_radius_m)
  movel([-0.080671, -0.870038, -2.777681, -1.064670, 1.570796, 1.490125],accel_mss,speed_ms,0,blend_radius_m)
  movel([-0.086258, -0.874029, -2.776840, -1.061520, 1.570796, 1.484538],accel_mss,speed_ms,0,blend_radius_m)
  movel([-0.091716, -0.878525, -2.775881, -1.057983, 1.570796, 1.479080],accel_mss,speed_ms,0,blend_radius_m)
  movel([-0.097048, -0.883450, -2.774817, -1.054122, 1.570796, 1.473748],accel_mss,speed_ms,0,blend_radius_m)
  movel([-0.102248, -0.888703, -2.773666, -1.050020, 1.570796, 1.468548],accel_mss,speed_ms,0,blend_radius_m)
  movel([-0.107307, -0.894193, -2.772444, -1.045751, 1.570796, 1.463490],accel_mss,speed_ms,0,blend_radius_m)
  movel([-0.112236, -0.899841, -2.771169, -1.041379, 1.570796, 1.458561],accel_mss,speed_ms,0,blend_radius_m)
  movel([-0.121695, -0.911274, -2.768525, -1.032590, 1.570796, 1.449101],accel_mss,speed_ms,0,blend_radius_m)
  movel([-0.123729, -0.913790, -2.767933, -1.030667, 1.570796, 1.447067],accel_mss,speed_ms,0,blend_radius_m)
  movel([-0.123869, -0.914204, -2.767835, -1.030351, 1.570796, 1.446928],accel_mss,speed_ms,0,blend_radius_m)
  movel([-0.123677, -0.914661, -2.767726, -1.030002, 1.570796, 1.447119],accel_mss,speed_ms,0,blend_radius_m)
  movel([-0.123269, -0.914995, -2.767647, -1.029747, 1.570796, 1.447527],accel_mss,speed_ms,0,blend_radius_m)
  speed_ms = 0.005
  movel([-0.123269, -0.905973, -2.761646, -1.044769, 1.570796, 1.447527],accel_mss,speed_ms,0,blend_radius_m)
  speed_ms = 0.040
  movel([-0.141809, -0.883593, -2.766751, -1.062045, 1.570796, 1.428988],accel_mss,speed_ms,0,blend_radius_m)
  speed_ms = 0.005
  movel([-0.141809, -0.892465, -2.772831, -1.047093, 1.570796, 1.428988],accel_mss,speed_ms,0,blend_radius_m)
  speed_ms = 0.025
  movel([-0.142140, -0.890069, -2.773363, -1.048956, 1.570796, 1.428656],accel_mss,speed_ms,0,blend_radius_m)
  movel([-0.142908, -0.888039, -2.773812, -1.050538, 1.570796, 1.427888],accel_mss,speed_ms,0,blend_radius_m)
  movel([-0.144096, -0.886428, -2.774166, -1.051795, 1.570796, 1.426701],accel_mss,speed_ms,0,blend_radius_m)
  movel([-0.145674, -0.885271, -2.774420, -1.052698, 1.570796, 1.425122],accel_mss,speed_ms,0,blend_radius_m)
  movel([-0.150413, -0.883591, -2.774786, -1.054012, 1.570796, 1.420383],accel_mss,speed_ms,0,blend_radius_m)
  movel([-0.151583, -0.882881, -2.774941, -1.054568, 1.570796, 1.419213],accel_mss,speed_ms,0,blend_radius_m)
  movel([-0.152432, -0.881952, -2.775142, -1.055295, 1.570796, 1.418365],accel_mss,speed_ms,0,blend_radius_m)
  movel([-0.152803, -0.880759, -2.775400, -1.056230, 1.570796, 1.417993],accel_mss,speed_ms,0,blend_radius_m)
  movel([-0.152536, -0.879243, -2.775727, -1.057419, 1.570796, 1.418260],accel_mss,speed_ms,0,blend_radius_m)
  movel([-0.151543, -0.877307, -2.776142, -1.058940, 1.570796, 1.419254],accel_mss,speed_ms,0,blend_radius_m)
  movel([-0.150265, -0.875802, -2.776463, -1.060124, 1.570796, 1.420531],accel_mss,speed_ms,0,blend_radius_m)
  movel([-0.148786, -0.874674, -2.776703, -1.061012, 1.570796, 1.422010],accel_mss,speed_ms,0,blend_radius_m)
  movel([-0.147199, -0.873874, -2.776873, -1.061643, 1.570796, 1.423597],accel_mss,speed_ms,0,blend_radius_m)
  movel([-0.144077, -0.873057, -2.777045, -1.062286, 1.570796, 1.426719],accel_mss,speed_ms,0,blend_radius_m)
  movel([-0.141608, -0.872929, -2.777072, -1.062388, 1.570796, 1.429189],accel_mss,speed_ms,0,blend_radius_m)
  movel([-0.142716, -0.870458, -2.777592, -1.064338, 1.570796, 1.428081],accel_mss,speed_ms,0,blend_radius_m)
  movel([-0.144331, -0.868590, -2.777983, -1.065816, 1.570796, 1.426465],accel_mss,speed_ms,0,blend_radius_m)
  movel([-0.148487, -0.865922, -2.778538, -1.067929, 1.570796, 1.422309],accel_mss,speed_ms,0,blend_radius_m)
  movel([-0.152861, -0.863396, -2.779059, -1.069934, 1.570796, 1.417935],accel_mss,speed_ms,0,blend_radius_m)
  movel([-0.154755, -0.861701, -2.779407, -1.071281, 1.570796, 1.416041],accel_mss,speed_ms,0,blend_radius_m)
  movel([-0.156241, -0.859450, -2.779866, -1.073072, 1.570796, 1.414555],accel_mss,speed_ms,0,blend_radius_m)
  movel([-0.156900, -0.857747, -2.780212, -1.074430, 1.570796, 1.413896],accel_mss,speed_ms,0,blend_radius_m)
  movel([-0.157213, -0.856169, -2.780530, -1.075689, 1.570796, 1.413584],accel_mss,speed_ms,0,blend_radius_m)
  movel([-0.157211, -0.854722, -2.780821, -1.076846, 1.570796, 1.413585],accel_mss,speed_ms,0,blend_radius_m)
  movel([-0.156924, -0.853413, -2.781083, -1.077893, 1.570796, 1.413873],accel_mss,speed_ms,0,blend_radius_m)
  movel([-0.156395, -0.852256, -2.781314, -1.078819, 1.570796, 1.414402],accel_mss,speed_ms,0,blend_radius_m)
  movel([-0.155651, -0.851246, -2.781515, -1.079628, 1.570796, 1.415145],accel_mss,speed_ms,0,blend_radius_m)
  movel([-0.154736, -0.850400, -2.781683, -1.080306, 1.570796, 1.416060],accel_mss,speed_ms,0,blend_radius_m)
  movel([-0.153677, -0.849722, -2.781817, -1.080850, 1.570796, 1.417119],accel_mss,speed_ms,0,blend_radius_m)
  movel([-0.152514, -0.849220, -2.781916, -1.081252, 1.570796, 1.418282],accel_mss,speed_ms,0,blend_radius_m)
  movel([-0.151289, -0.848907, -2.781978, -1.081504, 1.570796, 1.419507],accel_mss,speed_ms,0,blend_radius_m)
  movel([-0.148777, -0.848862, -2.781987, -1.081540, 1.570796, 1.422019],accel_mss,speed_ms,0,blend_radius_m)
  movel([-0.146432, -0.849641, -2.781833, -1.080915, 1.570796, 1.424365],accel_mss,speed_ms,0,blend_radius_m)
  movel([-0.144538, -0.851300, -2.781504, -1.079585, 1.570796, 1.426258],accel_mss,speed_ms,0,blend_radius_m)
  movel([-0.144291, -0.848272, -2.782103, -1.082014, 1.570796, 1.426505],accel_mss,speed_ms,0,blend_radius_m)
  movel([-0.144419, -0.845662, -2.782615, -1.084112, 1.570796, 1.426377],accel_mss,speed_ms,0,blend_radius_m)
  movel([-0.144844, -0.843379, -2.783060, -1.085950, 1.570796, 1.425952],accel_mss,speed_ms,0,blend_radius_m)
  movel([-0.147033, -0.837389, -2.784213, -1.090787, 1.570796, 1.423764],accel_mss,speed_ms,0,blend_radius_m)
  movel([-0.148397, -0.833034, -2.785038, -1.094317, 1.570796, 1.422399],accel_mss,speed_ms,0,blend_radius_m)
  movel([-0.148692, -0.831004, -2.785420, -1.095966, 1.570796, 1.422104],accel_mss,speed_ms,0,blend_radius_m)
  movel([-0.148704, -0.829055, -2.785784, -1.097551, 1.570796, 1.422092],accel_mss,speed_ms,0,blend_radius_m)
  movel([-0.148469, -0.827218, -2.786125, -1.099046, 1.570796, 1.422328],accel_mss,speed_ms,0,blend_radius_m)
  movel([-0.148012, -0.825514, -2.786439, -1.100435, 1.570796, 1.422784],accel_mss,speed_ms,0,blend_radius_m)
  movel([-0.147373, -0.823968, -2.786724, -1.101697, 1.570796, 1.423424],accel_mss,speed_ms,0,blend_radius_m)
  movel([-0.146578, -0.822600, -2.786974, -1.102814, 1.570796, 1.424218],accel_mss,speed_ms,0,blend_radius_m)
  movel([-0.145663, -0.821437, -2.787186, -1.103766, 1.570796, 1.425134],accel_mss,speed_ms,0,blend_radius_m)
  movel([-0.144659, -0.820504, -2.787356, -1.104530, 1.570796, 1.426137],accel_mss,speed_ms,0,blend_radius_m)
  movel([-0.143601, -0.819826, -2.787479, -1.105084, 1.570796, 1.427195],accel_mss,speed_ms,0,blend_radius_m)
  movel([-0.142525, -0.819426, -2.787551, -1.105412, 1.570796, 1.428271],accel_mss,speed_ms,0,blend_radius_m)
  movel([-0.141459, -0.819325, -2.787569, -1.105495, 1.570796, 1.429337],accel_mss,speed_ms,0,blend_radius_m)
  movel([-0.140438, -0.819552, -2.787528, -1.105308, 1.570796, 1.430358],accel_mss,speed_ms,0,blend_radius_m)
  movel([-0.139501, -0.820133, -2.787423, -1.104833, 1.570796, 1.431295],accel_mss,speed_ms,0,blend_radius_m)
  movel([-0.138678, -0.821086, -2.787250, -1.104053, 1.570796, 1.432119],accel_mss,speed_ms,0,blend_radius_m)
  movel([-0.138001, -0.822436, -2.787004, -1.102949, 1.570796, 1.432795],accel_mss,speed_ms,0,blend_radius_m)
  movel([-0.137501, -0.824198, -2.786682, -1.101510, 1.570796, 1.433296],accel_mss,speed_ms,0,blend_radius_m)
  movel([-0.136094, -0.820981, -2.787269, -1.104139, 1.570796, 1.434702],accel_mss,speed_ms,0,blend_radius_m)
  movel([-0.135009, -0.817887, -2.787829, -1.106673, 1.570796, 1.435788],accel_mss,speed_ms,0,blend_radius_m)
  movel([-0.134183, -0.814894, -2.788366, -1.109129, 1.570796, 1.436613],accel_mss,speed_ms,0,blend_radius_m)
  movel([-0.133548, -0.811973, -2.788885, -1.111531, 1.570796, 1.437248],accel_mss,speed_ms,0,blend_radius_m)
  movel([-0.131530, -0.800470, -2.790885, -1.121034, 1.570796, 1.439266],accel_mss,speed_ms,0,blend_radius_m)
  movel([-0.130668, -0.796155, -2.791618, -1.124617, 1.570796, 1.440128],accel_mss,speed_ms,0,blend_radius_m)
  movel([-0.129218, -0.790831, -2.792508, -1.129050, 1.570796, 1.441578],accel_mss,speed_ms,0,blend_radius_m)
  movel([-0.128102, -0.788113, -2.792957, -1.131319, 1.570796, 1.442695],accel_mss,speed_ms,0,blend_radius_m)
  movel([-0.126634, -0.785535, -2.793380, -1.133475, 1.570796, 1.444162],accel_mss,speed_ms,0,blend_radius_m)
  movel([-0.125742, -0.784337, -2.793575, -1.134478, 1.570796, 1.445055],accel_mss,speed_ms,0,blend_radius_m)
  movel([-0.123614, -0.782208, -2.793920, -1.136261, 1.570796, 1.447182],accel_mss,speed_ms,0,blend_radius_m)
  movel([-0.122358, -0.781316, -2.794063, -1.137009, 1.570796, 1.448438],accel_mss,speed_ms,0,blend_radius_m)
